(* IEC 61131-3 sources: daoli-st-library/DL_Device (part 36) *)

(* ---- FB_DL_VfdCapAgingEst.st ---- *)
(*
  ==================================================================
  组件名 Component  : FB_DL_VfdCapAgingEst
  分类   Category   : DL_Device
  前缀   Naming     : FB_DL_ ｜ b/n/u/f/t/e/st 类型前缀制（R265）
  码位   Code ID    : 16#0003_0725（故障级）｜ 16#0003_0726（信息级）
  版本   Version    : 1.0.0
  复杂度 Complexity  : 中
  功能   Purpose    : 母线电容老化趋势估计：纹波率实测值相对投运基线的长期比值监视
                      （电解电容容值衰减 → 纹波率单调爬升的运维预警）。
  开源溯源 Origin    : 公开公式 clean-room，参考公开电力电子运维工程口径的电解电容
                      纹波率基线比值判据（分类与公式借鉴，零代码复制），本件实现、
                      闸门与码位 100% 自有。
  许可证 License    : MIT
  参考   Reference  : IEC 61131-3:2013 §6.6 算术运算符；纹波率基线比值公开工程定义
  平台   Platform   : 纯 IEC 61131-3（四则 / 比较），三平台通用
  依赖   Depends    : 仅 Standard.library（无库调用、无定时器）
  分工声明 Split     : FB_DL_VfdDcBusRipple（瞬时纹波，R63 返修件）/ FB_DL_Brake
                      ResistorThermal（制动热）/ FB_DL_VfdThermalDerate（降额策略）
                      互引；本件为长期老化趋势，MANUAL 写明「瞬时监视与趋势估计
                      分层使用」（R216）。本件不实例依赖 VfdDcBusRipple，只收数值。
  归属 Ownership     : 本件无 TYPE 声明；全部引脚为 IEC 标准原生类型。
  ------------------------------------------------------------------
  边界 Boundary     :
                      一 组态闸结构早退（族② 判据，R1 同族教训出厂即正确）：
                         fRippleBasePct ≤ 0 或非有限（除子直穿防线）、fAgingLimPct ≤ 0
                         或非有限、fHystPct < 0 或非有限 → 组态码 0725 + 三件套 +
                         RETURN（除法段结构性不可达）；
                      二 fRipplePct 非有限或 < 0 → 该拍拒绝：比值冻结、迟滞态保持、
                         bValid = FALSE（丢弃 + 局部信息级计数，不外显 R62-D7 口径，
                         不影响趋势判据，禁污染物进除法）；
                      三 判据（带迟滞，两方向分别定义 R146）：fRippleRatioPct >
                         100 + fAgingLimPct 触发 bAgingHigh，回落 <
                         100 + fAgingLimPct×(1−fHystPct/100) 复原；
                      四 除子 fRippleBasePct > 0 已由段 2 结构早退证明（禁除零）；
                      五 负载可比性声明（写死）：本件假设同负载段比较，负载段切换时
                         调用方应 bEnable 短暂断开复位迟滞态——本件不自动判负载
                         （保持单一职责）；
                      六 bEnable = FALSE 的语义写死（FB33-4 声明行）：bAgingHigh 复位
                         + 比值冻结（运维趋势件，不丢历史）；
                      七 首拍 _bInit 全量初始化；无状态机（CASE N/A，R6 标注）；无
                         定时器 / 无边沿实例（段 0 无刷新对象）；无全局、无外部变量、
                         无物理地址、无指针。
  错误码 Codes      :
    16#0003_0725【故障级】组态非法（基线 ≤ 0 / 非有限；劣化阈值 ≤ 0 / 非有限；
                         迟滞 < 0 / 非有限）
    16#0003_0726【信息级】老化超限（bAgingHigh = TRUE，基线比超过 100 + 劣化阈值）
  码位反证 Note     :
    仅两码：0725 组态族为即刻判（与测点无关），0726 需比值已建立，处置人不同
    （组态工程师 / 运维），可由场景还原（R90）；fRipplePct 非有限拒绝拍不占码
    （bValid = FALSE 已足够表达，无额外处置信息，R90 不加码）。
  验收 Acceptance   :
    算法已证（脚本）：未跑 ｜ 编译器已证（三平台）：未跑
    V1 fRipplePct = fRippleBasePct → 比值 100%、bAgingHigh = FALSE
    V2 比值爬到 151%（限 150%）→ 触发；V3 回落 148%（迟滞未满足）→ 保持触发
    V4 回落 142% → 复原；V5 fRippleBasePct = 0 → 组态早退（R1 同族回归向量）
    V6 fRippleBasePct = NaN → 组态早退；V7 fRipplePct = NaN → 该拍拒绝不触发
    V8 fAgingLimPct = 0 → 组态早退（判据永假）
  修订记录 Revision  :
    2026-11-21  v1.0.0  R63 首版（批 4 · 序号 12）
  ==================================================================
*)
FUNCTION_BLOCK FB_DL_VfdCapAgingEst
VAR_INPUT
    bEnable       : BOOL := TRUE;  // 使能，FALSE 时判据复位 + 比值冻结（边界六）/ the enable, false resets the criterion and freezes the ratio
    fRipplePct    : LREAL := 0.0;  // 纹波率实测 [%]，由 FB_DL_VfdDcBusRipple 出口注入 / the measured ripple rate injected from the ripple monitor
    fRippleBasePct: LREAL := 5.0;  // 投运基线纹波率 [%]，须 > 0（除子）/ the commissioned baseline ripple rate, must be positive
    fAgingLimPct  : LREAL := 50.0; // 劣化阈值 [−]，相对基线百分比（50 即 150% 判劣化）/ the aging threshold relative to the baseline
    fHystPct      : LREAL := 5.0;  // 判据迟滞 [%]，须 ≥ 0 / the criterion hysteresis in percent, non negative
END_VAR
VAR_OUTPUT
    fRippleRatioPct : LREAL := 0.0;           // 基线比 fRipplePct/fRippleBasePct×100 [%] / the baseline ratio in percent
    bAgingHigh      : BOOL := FALSE;          // 老化超限判据（带迟滞）[-] / the aging high criterion with hysteresis
    bValid          : BOOL := FALSE;          // 判据可用 [-] / the criterion is usable
    eErr            : UDINT := 16#0000_0000;  // 错误码，0 = 正常 / the error code, zero is ok
    bError          : BOOL := FALSE;          // 故障标志（故障级码同拍置位，R45 配对）/ the fault flag raised with a fault level code
END_VAR
VAR
    _bInit      : BOOL := FALSE;   // 首拍初始化标志（R310 / FB50-2）/ the first scan flag
    _fRatio     : LREAL := 0.0;    // 基线比工作副本 [%] / the working baseline ratio
    _fRatioLast : LREAL := 0.0;    // 最近有效基线比（冻结源）[%] / the last valid ratio used while frozen
    _fTripLim   : LREAL := 0.0;    // 置警阈值 = 100 + 劣化阈值 [%] / the trip threshold
    _fReleLim   : LREAL := 0.0;    // 复原阈值 = 100 + 劣化阈值×(1−h) [%] / the release threshold
    _bAgingL    : BOOL := FALSE;   // 老化迟滞状态（跨拍保持）/ the aging hysteresis state
    _bFinBase   : BOOL := FALSE;   // 基线有限闸结果（逐拍重算）/ the baseline finiteness gate result
    _bFinLim    : BOOL := FALSE;   // 劣化阈值有限闸结果（逐拍重算）/ the threshold finiteness gate result
    _bFinHyst   : BOOL := FALSE;   // 迟滞有限闸结果（逐拍重算）/ the hysteresis finiteness gate result
    _bFinMeas   : BOOL := FALSE;   // 实测值有限闸结果（逐拍重算）/ the measurement finiteness gate result
    _bCfgBad    : BOOL := FALSE;   // 组态非法标记（逐拍重算）/ the configuration fault flag
    _nRejectCnt : DINT := 0;       // 实测值拒绝计数 [个]（仅局部留档，不外显，R62-D7 口径）/ the rejected measurement count, local only and never exposed
END_VAR  // R64 结构补齐：VAR 段缺失的 END_VAR（门禁机械修复）
VAR CONSTANT
    DL_VCA_PCT   : LREAL := 100.0; // 百分比换算与基线常量 [%] / the percentage scaling and the baseline constant
    DL_VCA_ZERO  : LREAL := 0.0;   // 实数零常量 [%] / the real zero constant
    DL_VCA_ONEI  : DINT := 1;      // 整型一常量 [个] / the integer one constant
    DL_VCA_ZEROI : DINT := 0;      // 整型零常量 [个] / the integer zero constant
END_VAR

// 段 0｜本件无定时器与边沿实例（纯趋势监视器，R6 标注 N/A），无刷新对象 / segment 0, no timers and no edge instances exist here

// 段 1｜首拍初始化（FB50-2）/ segment 1, the first scan init
IF NOT _bInit THEN // 首拍一拍 / the first scan
    _bInit := TRUE; // 置首拍标志 / raise the first scan flag
    _bAgingL := FALSE; // 迟滞态显式清零 / clear the hysteresis state explicitly
    _fRatioLast := DL_VCA_PCT; // 最近有效基线比显式预置 100%（首次有效计算前的安全占位）/ preset the last valid ratio to one hundred percent
    _nRejectCnt := DL_VCA_ZEROI; // 拒绝计数显式清零 [个] / clear the reject count explicitly
END_IF

// 段 2｜组态域闸结构早退（边界一，族② 判据：除子直穿防线先行，R272 全量点名）/ segment 2, the structural early exit on an illegal configuration
_bFinBase := (fRippleBasePct = fRippleBasePct) AND ((fRippleBasePct - fRippleBasePct) = (fRippleBasePct - fRippleBasePct)); // 基线有限 / the baseline is finite
_bFinLim := (fAgingLimPct = fAgingLimPct) AND ((fAgingLimPct - fAgingLimPct) = (fAgingLimPct - fAgingLimPct)); // 劣化阈值有限 / the threshold is finite
_bFinHyst := (fHystPct = fHystPct) AND ((fHystPct - fHystPct) = (fHystPct - fHystPct)); // 迟滞有限 / the hysteresis is finite
_bCfgBad := (NOT _bFinBase) OR (fRippleBasePct <= DL_VCA_ZERO)
         OR (NOT _bFinLim) OR (fAgingLimPct <= DL_VCA_ZERO)
         OR (NOT _bFinHyst) OR (fHystPct < DL_VCA_ZERO); // 组态非法 / an illegal configuration
IF _bCfgBad THEN // 组态非法：结构早退（出口三件套 + RETURN，除法段不可达）/ an illegal configuration exits structurally
    fRippleRatioPct := _fRatioLast; // 比值冻结最近有效值 [%]（禁自赋值出口，R261）/ freeze the last valid ratio
    bAgingHigh := FALSE; // 判据复位 / the criterion resets
    bValid := FALSE; // 判据不可用 / the criterion is not usable
    eErr := 16#0003_0725; // 故障级：组态非法 / fault grade, an illegal configuration
    bError := TRUE; // 同拍置故障标志（R45 配对）/ raise the fault flag on the same scan
    RETURN; // 结构早退 / the structural early exit
END_IF

// 段 3｜失能分支：判据复位 + 比值冻结（边界六声明行）/ segment 3, the disabled branch
IF NOT bEnable THEN // 失能 / disabled
    fRippleRatioPct := _fRatioLast; // 比值冻结最近有效值 [%]（运维趋势件，不丢历史）/ freeze the last valid ratio
    bAgingHigh := FALSE; // 判据复位 / the criterion resets
    bValid := FALSE; // 失能即不可用 / the criterion is not usable while disabled
    bError := FALSE; // 失能不是故障 / a disabled device is not a fault
    eErr := 16#0000_0000; // 失能不发码 / no code is emitted while disabled
    RETURN; // 早退 / early return
END_IF

// 段 4｜实测值拒绝闸（边界二：非有限或负值拒绝，禁污染物进除法）/ segment 4, the measurement rejection gate
_bFinMeas := (fRipplePct = fRipplePct) AND ((fRipplePct - fRipplePct) = (fRipplePct - fRipplePct)); // 实测值有限 / the measurement is finite
IF (NOT _bFinMeas) OR (fRipplePct < DL_VCA_ZERO) THEN // 实测坏或负值 / a broken or a negative measurement
    _nRejectCnt := _nRejectCnt + DL_VCA_ONEI; // 拒绝计数推进（仅局部留档，不外显）/ advance the reject count, local only
    fRippleRatioPct := _fRatioLast; // 比值冻结 [%] / freeze the ratio
    bAgingHigh := _bAgingL; // 迟滞态保持（拒绝拍不影响趋势判据）/ keep the hysteresis state
    bValid := FALSE; // 该拍不可用 / the scan is not usable
    eErr := 16#0000_0000; // 拒绝拍不发码（bValid = FALSE 已足够表达，R90 不加码）/ no code for a rejected scan
    bError := FALSE; // 无故障 / no fault
    RETURN; // 早退，除法不可达 / early return, the division is unreachable
END_IF

// 段 5｜基线比计算（除子 fRippleBasePct > 0 已由段 2 证明，禁除零）/ segment 5, the baseline ratio computation
_fRatio := (fRipplePct / fRippleBasePct) * DL_VCA_PCT; // 基线比 [%]，除子已证 > 0 / the baseline ratio with the proven divisor
_fRatioLast := _fRatio; // 最近有效基线比快照 [%] / snapshot the valid ratio
_fTripLim := DL_VCA_PCT + fAgingLimPct; // 置警阈值 [%] / the trip threshold
_fReleLim := DL_VCA_PCT + (fAgingLimPct * ((DL_VCA_PCT - fHystPct) / DL_VCA_PCT)); // 复原阈值 [%] / the release threshold

// 段 6｜老化判据迟滞（边界三，两方向分别定义，R146）/ segment 6, the aging hysteresis
IF NOT _bAgingL THEN // 未报警态 / the released state
    IF _fRatio > _fTripLim THEN // 超过置警阈值 / above the trip threshold
        _bAgingL := TRUE; // 置迟滞状态 / set the hysteresis state
    END_IF
ELSE // 已报警态 / the tripped state
    IF _fRatio < _fReleLim THEN // 回落低于复原阈值 / below the release threshold
        _bAgingL := FALSE; // 复原 / release
    END_IF
END_IF

// 段 7｜统一出口（迟滞状态派生，R187 / FB51-8）/ segment 7, the unified outlet
fRippleRatioPct := _fRatio; // 基线比出口 [%] / the ratio outlet
bAgingHigh := _bAgingL; // 判据出口 / the criterion outlet
bValid := TRUE; // 判据可用 / the criterion is usable
bError := FALSE; // 无故障 / no fault
IF _bAgingL THEN // 老化超限（信息级）/ the aging is high, informational
    eErr := 16#0003_0726; // 信息级：基线比超过 100 + 劣化阈值 / informational, the ratio exceeds the aging threshold
ELSE // 无事件 / no event
    eErr := 16#0000_0000; // 正常 / ok
END_IF
END_FUNCTION_BLOCK

(* ---- FB_DL_VfdCtrlWordBuild.st ---- *)
(*
  道莅工业代码库 | DL_Device | FB_DL_VfdCtrlWordBuild
  版本: 1.0.0 | 日期: 2026-11-23 | 轮次: R75
  开源溯源: brOscatLib (github.com/brOscatLib) / MIT / 借鉴 CtrlWordBuild 的语义，代码为 clean-room 重写
  功能: 变频器控制字编码——目标状态号（bit0..3）+ 命令位（运行/自由停车/直流
        制动/快速停止/反转/复位脉冲）按固定位图组装控制字；与 FB_DL_VfdStateWordMatch
        成对（编码/判码）。变换型 FB：无相位机，每拍独立全量重算。
  兼容性: CODESYS 3.5 / TwinCAT 3 / 汇川 InoProShop；仅依赖标准 R_TRIG，零厂商私有库
  接口: 输入 bEn/uStateNo（0..15，越界钳 15 并置信息码）/六命令位；输出
        wCtrlWord/uStateEff（钳位后状态号）/bRangeInfo/bError/nErrId。
  位图定义（bit0..3 = 目标状态号，与 C04 判码件低 4 位状态号口径一致）:
    bit4 = 运行命令 bRunCmd            bit5 = 非自由停车（1=斜坡停车可用）
    bit6 = 直流制动 bDCBrake           bit7 = 复位脉冲（R_TRIG 单拍）
    bit11 = 反转 bReverse              bit13 = 快速停止 bQuickStop
  码表: 16#0003_040F 信息级：目标状态号越域钳 15（每拍重算，非锁存）
        码段说明：0003 段信息子带 04xx，槽位经全库实扫空闲。
  边界: ① uStateNo > 15 → 钳 15 + bRangeInfo（本件无故障级路径，bError 恒 FALSE）；
        ② bit7 复位脉冲由 R_TRIG 单拍化（不复位脉冲不驻留控制字）；
        ③ bEn = FALSE 时控制字输出 16#0000（全零安全侧）；
        ④ R_TRIG 段 0 无条件周期刷新；⑤ 零全局耦合。
  邻件比对: StatusWordSegDecoder（通用分段译码 vs 本件变频器控制字编码组装）。
  修订历史: 2026-11-23 v1.0.0 R75 首版（复杂件批 B2 · C10）
*)

FUNCTION_BLOCK FB_DL_VfdCtrlWordBuild
VAR_INPUT
    bEn         : BOOL := FALSE;    // 编码使能（FALSE 输出全零控制字）[-] | Build enable, FALSE outputs zero word
    uStateNo    : UINT := 0;        // 目标状态号，域 [0, 15]，越界钳 15 [号] | Target state number, clamped to 15
    bRunCmd     : BOOL := FALSE;    // 运行命令（bit4）[-] | Run command bit
    bCoastStop  : BOOL := FALSE;    // 自由停车选择（TRUE 时 bit5=0）[-] | Coast stop select, TRUE clears bit5
    bDCBrake    : BOOL := FALSE;    // 直流制动（bit6）[-] | DC brake bit
    bQuickStop  : BOOL := FALSE;    // 快速停止（bit13）[-] | Quick stop bit
    bReverse    : BOOL := FALSE;    // 反转（bit11）[-] | Reverse bit
    bResetCmd   : BOOL := FALSE;    // 故障复位命令（bit7，沿触发单拍）[-] | Fault reset command, edge one-shot
END_VAR
VAR_OUTPUT
    wCtrlWord  : WORD;              // 组装控制字出口（bEn=FALSE 时全零）[-] | Built control word outlet
    uStateEff  : UINT;              // 钳位后状态号出口 [号] | Clamped state number outlet
    bRangeInfo : BOOL;              // 状态号越域钳位当拍信息 [-] | Range clamp info this scan
    bError     : BOOL;              // 故障标志（本件无故障路径，恒 FALSE）[-] | Error flag, no fault paths
    nErrId     : UDINT;             // 事件码，0 = 无事件 | Event code, 0 = none
END_VAR
VAR
    _uStateEff : UINT := 0;         // 钳位状态号内部镜像 [号] | Clamped state number mirror
    _wOut      : WORD := 16#0000;   // 组装暂存字 [-] | Build staging word
    _bRange    : BOOL;              // 越域当拍量 [-] | Range violation this scan
    rtResetCmd : R_TRIG;            // 复位脉冲沿实例，段 0 无条件刷新 | Reset pulse edge instance
END_VAR

(* —— 段 0：沿实例无条件周期刷新（R7 红线） —— *)
rtResetCmd(CLK := bResetCmd);                 // 复位脉冲沿每拍必调 / Reset pulse edge every scan

(* —— 段 1：状态号钳位（越域置当拍信息量） —— *)
_uStateEff := uStateNo;                       // 状态号暂存 / State number staging
_bRange := FALSE;                             // 越域当拍量预清 / Range flag preset
IF _uStateEff > 15 THEN
    _uStateEff := 15;                         // 越域钳 15 / Clamp to 15
    _bRange := TRUE;                          // 置越域信息量 / Set range info
END_IF

(* —— 段 2：控制字位图组装（bit0..3 状态号） —— *)
_wOut := INT_TO_WORD(UINT_TO_INT(_uStateEff)) AND 16#000F;    // 状态号入低 4 位（掩码兜底）/ State number to low nibble
IF bRunCmd THEN
    _wOut := _wOut OR 16#0010;                // bit4 运行命令 / Run command bit
END_IF
IF NOT bCoastStop THEN
    _wOut := _wOut OR 16#0020;                // bit5 斜坡停车可用（非自由停车）/ Ramp stop available bit
END_IF
IF bDCBrake THEN
    _wOut := _wOut OR 16#0040;                // bit6 直流制动 / DC brake bit
END_IF
IF rtResetCmd.Q THEN
    _wOut := _wOut OR 16#0080;                // bit7 复位脉冲（仅沿当拍驻留）/ Reset pulse bit, one scan only
END_IF
IF bReverse THEN
    _wOut := _wOut OR 16#0800;                // bit11 反转 / Reverse bit
END_IF
IF bQuickStop THEN
    _wOut := _wOut OR 16#2000;                // bit13 快速停止 / Quick stop bit
END_IF

(* —— 段 3：出口单点映射（名实同源；信息码每拍重算） —— *)
IF bEn THEN
    wCtrlWord := _wOut;                       // 使能输出组装字 / Enabled, output built word
ELSE
    wCtrlWord := 16#0000;                     // 未使能输出全零（安全侧） / Disabled, output zero word
END_IF
uStateEff := _uStateEff;                      // 钳位状态号出口 / Clamped state outlet
bRangeInfo := _bRange;                        // 越域信息出口 / Range info outlet
bError := FALSE;                              // 本件无故障级路径（头注释声明）/ No fault paths by design
IF _bRange THEN
    nErrId := 16#0003_040F;                   // 信息级：状态号越域钳位 / Info: state number clamped
ELSE
    nErrId := 16#0000_0000;                   // 无事件 / No event
END_IF

END_FUNCTION_BLOCK

(* ---- FB_DL_VfdGeneric.st ---- *)
(*==============================================================================
 * 组件名称 (Component)  : FB_DL_VfdGeneric
 * 所属子库 (Sublibrary) : DL_Device
 * 当前版本 (Version)    : 1.0.1
 * 兼容性   (Platform)   : CODESYS 3.5 / TwinCAT 3 / 汇川 InoProShop / Machine Expert
 *                         仅依赖 Standard.library（TON / R_TRIG / TP），零厂商方言
 * 分类     (Category)   : 设备执行器功能块（Function Block，实现 I_DL_VfdDrive）
 * 功能简述 (Function)   : 通用变频器端子型控制功能块。正/反转端子互斥
 *                         （出口断言 + 冲突安全侧停止）、点动优先覆盖运行、
 *                         多段速表/模拟量给定双通道频率设定（越界钳位）、
 *                         频率给定模拟量域线性映射、指令-反馈校验窗、驱动
 *                         故障锁存与复位端子定宽脉冲重试；状态机
 *                         E_DL_VfdState + CASE + ELSE 兜底。
 * 接口实现 (Implements) : I_DL_VfdDrive。接口 OUT 列同名成员（eState/
 *                         fFreqSetpoint/fFreqActual/bRunning/bFault/
 *                         uErrorId）按 R22 以只读 PROPERTY GET 承载（内部
 *                         镜像同源），非接口成员 bRunFwdOut/bRunRevOut/
 *                         bJogOut/bFaultResetOut/fFreqRefPercent/uPresetCode
 *                         保留 VAR_OUTPUT；方法 CmdRun/CmdStop/CmdJog/
 *                         SetFrequency/SelectPresetSpeed/CmdReset 全部在
 *                         本文件尾部落地。
 * 开源溯源 (Origin)     : 来源标签 lbp-basic-process / lbp-device
 *                         （RAW_NOTES_R6 S-1 + S-4：变频器端子标准信号集
 *                         ——正反转互斥、点动优先、多段速 DI 组合、模拟
 *                         量频率给定线性映射、故障复位端子脉冲等行业公知
 *                         工程惯例，公开技术资料，仅借鉴通用信号域语义；
 *                         状态机、钳位与互斥实现、故障码按本库红线独立
 *                         设计，clean-room 未复制源码）。
 * 红线自检 (Redline)    : R1 零全局变量表/外部变量引用 ✓｜R2 零物理 IO 地址 ✓
 *                         R3 纯 IEC 61131-3 ✓｜R4 防除零/防越界/非有限值
 *                         防御/浮点容差比较 ✓｜R5 全变量中英双语同行注释 ✓
 *                         R6 ENUM+CASE+ELSE ✓｜R7 三个定时器/边缘/脉冲实例
 *                         主体最前部无条件刷新 ✓
 * 公约遵循 (Convention) : 0.1/R23 本块为纯事件型状态机（BOOL 指令/反馈 +
 *                         频率标量直通计算，无积分/滤波类连续量同步语义），
 *                         免首扫，无内部初始化标志。
 *                         0.7 故障码段位 16#0003_xxxx：【故障级】0003_0250
 *                         驱动故障 / 0003_0251 启动反馈超时 / 0003_0252
 *                         非法状态，R15 锁存仅复位脉冲路径可清；【信息级】
 *                         0003_0106 正反转指令冲突 / 0003_0107 频率设定
 *                         钳位/段速选择越界（瞬时型每拍重算，0.15）。
 * 偏离留档 (Deviation)  : 依 R11 头注释留档，共 2 条：
 *                         ① 信息级码：规格原分配 0003_0103/0104，经与子库
 *                           VERSION.md 故障码表核对，R5 已占用 0102~0104
 *                           （AnalogTransmitter），依公约 0.7 冲突顺延为
 *                           0003_0106/0107（0105 经终审裁定空置：重启抑制
 *                           拒绝统一沿用 DolMotor 既有语义码位 0003_0208，
 *                           见 FB_DL_StarDeltaMotor 终审记录）。
 *                         ② 点动频率：规格设计要点"点动频率取 aPresetFreq[1]
 *                           （注释声明）"落为引脚注释声明——本块不因点动切
 *                           换频率通道（端子型变频器点动频率由驱动器内部组
 *                           态承担），段速 1 兼作点动频率域供现场整定选用。
 * 修订历史 (Revision)   :
 *   2026-11-15  v1.0.0  首版入库（R6 轮 · DL_Device 阀门/驱动族深化）
 *   2026-11-15  v1.0.1  终审修复【致命】复位端子脉冲触发时序：原实现
 *                       _bResetPulseReq 于主体末尾同拍自清，TP 实例（段 1
 *                       最前部刷新）永远采不到 TRUE 入参，bFaultResetOut
 *                       恒 FALSE，故障复位端子脉冲永不输出（验收向量 V5
 *                       不成立，R13 逐拍推演复现）。修法：自清动作移至
 *                       TP 实例调用之后。另补点动频率引脚注释声明（R11
 *                       偏离②）。引脚契约零变更。
 *============================================================================*)
FUNCTION_BLOCK FB_DL_VfdGeneric IMPLEMENTS I_DL_VfdDrive
VAR_INPUT
    bDriveEnable     : BOOL;            // 驱动使能/上电（Drive enable），FALSE → 未使能态全部输出切断 / Drive enable, FALSE cuts off all outputs
    bCmdRunFwd       : BOOL;            // 正转运行指令（Run forward command），电平生效 / Run forward command, level effective
    bCmdRunRev       : BOOL;            // 反转运行指令（Run reverse command），电平生效；与正转同拍为真 → 冲突安全侧停止 / Run reverse command, conflict with forward stops safely
    bCmdJogFwd       : BOOL;            // 正向点动指令（Jog forward command），电平生效，优先级高于运行指令；点动频率不在本块内切换通道——端子型惯例由驱动器内部点动频率组态承担，亦可现场将 aPresetFreq[1] 整定为点动频率域（段速 1 兼作点动频率） / Jog forward command, level effective, priority over run; jog frequency not switched by this block, use drive-internal jog frequency or tune aPresetFreq[1] as the jog frequency domain
    bFbRunning       : BOOL;            // 运行反馈（Running feedback），TRUE=驱动输出运行中 / Running feedback, TRUE = drive output running
    bFbFault         : BOOL;            // 驱动故障反馈（Drive fault feedback），TRUE=故障 / Drive fault feedback, TRUE = faulty
    bFbAtSpeed       : BOOL;            // 频率到达反馈（At-speed feedback），TRUE=输出频率到达设定容差带 / At-speed feedback, TRUE = output frequency reached setpoint band
    fFreqCmd         : REAL;            // 频率设定（Frequency command）[Hz]，0..fFreqMax，越界钳位信息级 / Frequency command [Hz], clamped with info code
    fFreqActual      : REAL;            // 频率反馈（Frequency feedback）[Hz]，非有限值防御 / Frequency feedback [Hz], non-finite defended
    aPresetFreq      : ARRAY[1..7] OF REAL; // 多段速频率表（Preset speed table）[Hz]，段速值由现场整定注入 / Preset speed table [Hz], field-tuned values injected
    nPresetSel       : USINT;           // 段速选择（Preset speed select），0=模拟量给定、1..7=段速，越界按 0 处理并置码 / Preset select, 0 = analog reference, 1..7 = steps, out-of-range treated as 0 with code
    fFreqMax         : REAL := 50.0;    // 频率上限（Max frequency）[Hz]，默认 50.0 / Maximum frequency [Hz], default 50.0
    tFbWindow        : TIME := T#1S;    // 指令-反馈校验窗口（Feedback check window），T#0S=免校验 / Feedback check window, T#0S disables the check
    tFaultResetPulse : TIME := T#500MS; // 故障复位脉冲宽度（Fault reset pulse）/ Fault reset pulse width
    bReset           : BOOL;            // 故障复位请求（Fault reset request），上升沿生效 / Fault reset request, rising edge effective
END_VAR

VAR_OUTPUT
    bRunFwdOut      : BOOL;             // 正转端子输出（Run forward terminal）/ Run forward terminal output
    bRunRevOut      : BOOL;             // 反转端子输出（Run reverse terminal）/ Run reverse terminal output
    bJogOut         : BOOL;             // 点动端子输出（Jog terminal）/ Jog terminal output
    bFaultResetOut  : BOOL;             // 故障复位端子输出（Fault reset terminal），tFaultResetPulse 定宽单发 / Fault reset terminal, one-shot fixed-width pulse
    fFreqRefPercent : REAL;             // 频率给定模拟量输出（Frequency reference analog out）[%]，0~100 线性映射 fFreqMax / Analog frequency reference [%], linear over fFreqMax
    uPresetCode     : USINT;            // 段速选择码输出（Preset speed code），映射 DI 多段速端子组合 0..7 / Preset speed code mapped to DI terminal group 0..7
END_VAR

VAR
    _eState         : E_DL_VfdState := E_DL_VfdState.eDisabled; // 内部状态机步序（Internal state step），外部经属性只读 / Internal state, read-only via property
    _bFaultLatch    : BOOL;             // 故障锁存标志（Fault latch flag），仅复位脉冲路径清除 / Fault latch flag, cleared only via reset pulse path
    _uErrorIdInt    : UDINT;            // 内部故障码寄存（Internal error register），故障级与信息级共用 / Internal error register, fault and info codes share it
    _uInfoCode      : UDINT;            // 本拍信息级码（Info code this cycle），瞬时型每拍重算（0.15）/ Transient info code recomputed each cycle
    _bPendRunFwd    : BOOL;             // 方法正转保持锁存（Method run-forward hold latch）/ Method run-forward hold latch
    _bPendRunRev    : BOOL;             // 方法反转保持锁存（Method run-reverse hold latch）/ Method run-reverse hold latch
    _bJogHold       : BOOL;             // 方法点动保持锁存（Method jog hold latch）/ Method jog hold latch
    _bPendReset     : BOOL;             // 方法复位请求（Method reset request）/ Method reset request
    _bResetPulseReq : BOOL;             // 复位脉冲单拍触发请求（Reset pulse trigger request），置位一拍 / One-cycle reset pulse trigger request
    _fFreqMethodVal : REAL;             // 方法频率设定值（Method frequency value）[Hz] / Frequency value set via method
    _bFreqMethodAct : BOOL;             // 方法频率设定激活（Method frequency active），激活后覆盖引脚给定 / Method frequency active, overrides pin reference
    _uPresetMethod  : USINT;            // 方法段速选择值（Method preset select value）/ Preset select value set via method
    _bPresetMethodAct : BOOL;           // 方法段速选择激活（Method preset select active）/ Method preset select active flag
    _fFreqMaxEff    : REAL := 50.0;     // 防御后频率上限（Sanitized max frequency）[Hz] / Sanitized maximum frequency
    _fFreqCmdEff    : REAL := 0.0;      // 防御后模拟量给定（Sanitized analog command）[Hz]，非数回零 / Sanitized analog command, NaN falls back to zero
    _fFreqSetInt    : REAL := 0.0;      // 钳位后生效频率设定（Effective clamped setpoint）[Hz] / Effective clamped frequency setpoint
    _fFreqActHold   : REAL := 0.0;      // 末次有效频率反馈（Last valid frequency feedback）[Hz] / Last valid frequency feedback hold carrier
    _uPresetSelEff  : USINT;            // 钳位后生效段速选择（Effective clamped preset select），0..7 / Effective preset select clamped to 0..7
    _bRunFwd        : BOOL;             // 合成正转指令（Merged run-forward command），引脚 OR 方法锁存 / Merged forward command, pin OR method latch
    _bRunRev        : BOOL;             // 合成反转指令（Merged run-reverse command），引脚 OR 方法锁存 / Merged reverse command, pin OR method latch
    _bJog           : BOOL;             // 合成点动指令（Merged jog command），引脚 OR 方法锁存 / Merged jog command, pin OR method latch
    _bConflict      : BOOL;             // 正反转同拍冲突（Forward/reverse conflict this cycle）/ Forward-reverse conflict flag
    _bFbWinEn       : BOOL;             // 反馈校验窗使能（Feedback window enable），窗口参数大于零有效 / Feedback window enable, active when window above zero
    _bInFbWin       : BOOL;             // 反馈校验窗计时条件（Feedback window timing condition）/ Timing condition of feedback window
    _fbTrigReset    : R_TRIG;           // 引脚复位上升沿（Pin reset edge）/ Pin reset rising edge
    _fbTonFbWindow  : TON;              // 启动反馈校验窗定时器（Startup feedback window timer）/ Startup feedback window timer
    _fbTpResetPulse : TP;               // 复位端子定宽脉冲定时器（Reset terminal pulse timer），IEC 标准 TP / Reset terminal pulse timer, IEC standard TP
END_VAR

METHOD CmdRun : BOOL
VAR_INPUT
    bFwd : BOOL; // 方向选择（Direction select），TRUE=正转 / FALSE=反转 / TRUE = forward, FALSE = reverse
END_VAR
IF _bFaultLatch OR (_eState = E_DL_VfdState.eFault) OR (_eState = E_DL_VfdState.eDisabled) THEN
    CmdRun := FALSE;          // 故障/未使能态拒绝（Rejected in fault or disabled state）
ELSE
    IF bFwd THEN
        _bPendRunFwd := TRUE; // 登记正转保持锁存（Register forward hold latch）
        _bPendRunRev := FALSE; // 互斥注销反转锁存（Cancel opposite latch）
    ELSE
        _bPendRunRev := TRUE; // 登记反转保持锁存（Register reverse hold latch）
        _bPendRunFwd := FALSE; // 互斥注销正转锁存（Cancel opposite latch）
    END_IF
    CmdRun := TRUE;           // 受理成功（Accepted）
END_IF

(*------------------------------------------------------------------------------
 * 方法: CmdStop —— 停止指令：撤销运行/点动锁存，无条件受理。
 *      Method CmdStop - revokes run and jog latches, unconditionally accepted.
 *------------------------------------------------------------------------------*)
    END_METHOD

METHOD CmdStop : BOOL
VAR_INPUT
END_VAR
_bPendRunFwd := FALSE;        // 撤销正转锁存（Release forward latch）
_bPendRunRev := FALSE;        // 撤销反转锁存（Release reverse latch）
_bJogHold    := FALSE;        // 撤销点动保持（Release jog hold）
CmdStop := TRUE;              // 无条件受理（Unconditionally accepted）

(*------------------------------------------------------------------------------
 * 方法: CmdJog —— 点动指令（bFwd=TRUE 登记保持 / FALSE 撤销）。故障态拒绝。
 *      Method CmdJog - jog hold register/release, rejected in fault state.
 *------------------------------------------------------------------------------*)
    END_METHOD

METHOD CmdJog : BOOL
VAR_INPUT
    bFwd : BOOL; // 点动方向（Jog direction），TRUE=正向登记 / FALSE=撤销保持 / TRUE = register, FALSE = release
END_VAR
IF _bFaultLatch OR (_eState = E_DL_VfdState.eFault) THEN
    CmdJog := FALSE;          // 故障态拒绝（Rejected in fault state）
ELSE
    _bJogHold := bFwd;        // 登记或撤销点动保持（Register or release jog hold）
    CmdJog := TRUE;           // 受理成功（Accepted）
END_IF

(*------------------------------------------------------------------------------
 * 方法: SetFrequency —— 频率设定 [Hz]，越界/非有限值拒绝返回 FALSE。
 *      Method SetFrequency - frequency set, out-of-range or NaN returns FALSE.
 *------------------------------------------------------------------------------*)
    END_METHOD

METHOD SetFrequency : BOOL
VAR_INPUT
    fHz : REAL; // 频率设定值（Frequency value）[Hz]，域 0..fFreqMax / Frequency value [Hz], range 0..fFreqMax
END_VAR
IF (fHz <> fHz) OR (fHz < 0.0) OR (fHz > _fFreqMaxEff) THEN
    SetFrequency := FALSE;    // 非数或越域拒绝（Rejected on NaN or out of range）
ELSE
    _fFreqMethodVal := fHz;   // 登记方法频率设定（Register method frequency value）
    _bFreqMethodAct := TRUE;  // 激活方法给定通道（Activate method reference channel）
    SetFrequency := TRUE;     // 受理成功（Accepted）
END_IF

(*------------------------------------------------------------------------------
 * 方法: SelectPresetSpeed —— 多段速选择，0=模拟量给定、1..7=段速，越界拒绝。
 *      Method SelectPresetSpeed - preset select, 0 = analog, 1..7 = steps.
 *------------------------------------------------------------------------------*)
    END_METHOD

METHOD SelectPresetSpeed : BOOL
VAR_INPUT
    nIdx : USINT; // 段速索引（Preset index），0=模拟量给定 / 1..7=段速 / Preset index, 0 = analog reference, 1..7 = steps
END_VAR
IF nIdx <= 7 THEN
    _uPresetMethod := nIdx;   // 登记方法段速选择（Register method preset value）
    _bPresetMethodAct := TRUE; // 激活方法段速通道（Activate method preset channel）
    SelectPresetSpeed := TRUE; // 受理成功（Accepted）
ELSE
    SelectPresetSpeed := FALSE; // 越界拒绝（Rejected on out-of-range index）
END_IF

(*------------------------------------------------------------------------------
 * 方法: CmdReset —— 复位指令，返回是否受理（存在锁存故障时为 TRUE）。
 *      Method CmdReset - reset command, returns TRUE only when latch exists.
 *------------------------------------------------------------------------------*)
    END_METHOD

METHOD CmdReset : BOOL
VAR_INPUT
END_VAR
IF _bFaultLatch OR (_eState = E_DL_VfdState.eFault) THEN
    _bPendReset := TRUE;      // 登记复位请求，主体状态机消化（Register reset request, consumed by body）
    CmdReset := TRUE;         // 可复位（Resettable）
ELSE
    CmdReset := FALSE;        // 无故障可复位（Nothing to reset）
END_IF

(*------------------------------------------------------------------------------
 * 属性: eState（GET）—— 当前状态机状态只读视图。
 *      Property eState (GET) - read-only view of the current state machine state.
 *------------------------------------------------------------------------------*)
    END_METHOD

// ============================================================================
// 段 1｜定时器与边缘检测实例无条件周期刷新（R7：严禁置于 IF/CASE 分支内）
//      Unconditional per-cycle refresh of all timer and edge instances (R7)
// ============================================================================
_fbTrigReset(CLK := bReset);
_bFbWinEn := (tFbWindow > T#0S);      // 窗口为零 = 免校验（Zero window = check disabled）
_bInFbWin := ((_eState = E_DL_VfdState.eRunningFwd) OR (_eState = E_DL_VfdState.eRunningRev))
             AND (NOT bFbRunning) AND _bFbWinEn; // 运行态且反馈未到才计时（Timing only while running and feedback pending）
_fbTonFbWindow(IN := _bInFbWin, PT := tFbWindow);
_fbTpResetPulse(IN := _bResetPulseReq, PT := tFaultResetPulse); // 复位端子定宽脉冲（Fixed-width reset terminal pulse）
_bResetPulseReq := FALSE;             // 单拍触发请求在 TP 采样后立即自清：TP 于本拍见到
                                      // TRUE 并起振，下一拍入参回落 FALSE，定宽由 TP 保持
                                      // （One-cycle trigger cleared right after TP sampling）

// ============================================================================
// 段 2｜参数防御（0.8：非数自比检测，默认值先赋）+ 指令合成与钳位
//      Parameter sanitation (0.8 NaN self-compare) + command merge and clamping
// ============================================================================
_uInfoCode := 0;                      // 本拍信息级码先归零，事件段重算（Info code preset zero, recomputed in event chain）
_fFreqMaxEff := fFreqMax;             // 频率上限镜像（Max frequency mirror）
IF _fFreqMaxEff <> _fFreqMaxEff THEN  // 非数自比检测（NaN self-compare test）
    _fFreqMaxEff := 50.0;             // 回落默认上限（Fallback to default max）
END_IF
IF ABS(_fFreqMaxEff) < 1E-6 THEN
    _fFreqMaxEff := 1E-6;             // 防除零：上限退化时钳最小正值（Divide-by-zero guard, degenerate max clamped to tiny positive）
END_IF

IF _bFreqMethodAct THEN
    _fFreqCmdEff := _fFreqMethodVal;  // 方法设定覆盖引脚给定（Method value overrides pin reference）
ELSE
    _fFreqCmdEff := fFreqCmd;         // 引脚模拟量给定（Pin analog reference）
END_IF
IF _fFreqCmdEff <> _fFreqCmdEff THEN  // 非数自比检测（NaN self-compare test）
    _fFreqCmdEff := 0.0;              // 非数给定回零（NaN reference falls back to zero）
END_IF
IF _fFreqCmdEff < 0.0 THEN
    _fFreqCmdEff := 0.0;              // 负给定下限钳位（Negative reference clamped to zero）
    _uInfoCode := 16#0003_0107;       // 0003_0107 频率设定钳位【信息级】/ Frequency clamped, info level
END_IF
IF _fFreqCmdEff > _fFreqMaxEff THEN
    _fFreqCmdEff := _fFreqMaxEff;     // 超上限钳位（Reference clamped to max）
    _uInfoCode := 16#0003_0107;       // 0003_0107 频率设定钳位【信息级】/ Frequency clamped, info level
END_IF

IF fFreqActual = fFreqActual THEN     // 频率反馈有效性（Frequency feedback validity）
    _fFreqActHold := fFreqActual;     // 更新末次有效反馈（Update last valid feedback）
END_IF                                 // 非有限值保持末次有效值（Non-finite holds last valid）

// 段速选择钳位：越界按 0 处理并置码（Preset select clamped, out-of-range as 0 with code）
IF _bPresetMethodAct THEN
    _uPresetSelEff := _uPresetMethod; // 方法段速选择覆盖引脚（Method preset overrides pin）
ELSIF nPresetSel <= 7 THEN
    _uPresetSelEff := nPresetSel;     // 引脚段速选择合法（Pin preset select valid）
ELSE
    _uPresetSelEff := 0;              // 越界按模拟量给定处理（Out-of-range treated as analog reference）
    _uInfoCode := 16#0003_0107;       // 0003_0107 段速选择越界【信息级】/ Preset select out of range, info level
END_IF

// 生效频率设定：段速优先，模拟量给定兜底（Effective setpoint: preset first, analog fallback）
IF (_uPresetSelEff >= 1) AND (_uPresetSelEff <= 7) THEN
    _fFreqSetInt := aPresetFreq[_uPresetSelEff];       // 取段速表值（Take preset table value, index proven 1..7）
    IF _fFreqSetInt <> _fFreqSetInt THEN
        _fFreqSetInt := 0.0;                           // 段速值非数回零防御（NaN preset falls back to zero）
    END_IF
ELSE
    _fFreqSetInt := _fFreqCmdEff;     // 模拟量给定通道（Analog reference channel）
END_IF

// 指令合成与冲突判定（Command merge and conflict evaluation）
_bRunFwd := bCmdRunFwd OR _bPendRunFwd; // 合成正转（Merged forward）
_bRunRev := bCmdRunRev OR _bPendRunRev; // 合成反转（Merged reverse）
_bJog := bCmdJogFwd OR _bJogHold;       // 合成点动，优先级最高（Merged jog, highest priority）
_bConflict := _bRunFwd AND _bRunRev;    // 同拍正反转冲突（Same-cycle conflict）
IF _bConflict THEN
    _uInfoCode := 16#0003_0106;         // 0003_0106 正反转指令冲突【信息级】/ Forward-reverse conflict, info level
END_IF

// ============================================================================
// 段 3｜驱动故障全局监视（优先级最高）：故障反馈置锁存
//      Drive fault global monitor (highest priority): fault feedback latches
// ============================================================================
IF bFbFault THEN
    _bFaultLatch := TRUE;               // 驱动故障锁存（Drive fault latch）
    _uErrorIdInt := 16#0003_0250;       // 0003_0250 驱动故障【故障级】/ Drive fault, fault level
    _eState      := E_DL_VfdState.eFault; // 强制故障态（Force fault state）
ELSIF (_eState = E_DL_VfdState.eRunningFwd) OR (_eState = E_DL_VfdState.eRunningRev) THEN
    IF _bFbWinEn AND _fbTonFbWindow.Q AND (NOT bFbRunning) THEN
        _bFaultLatch := TRUE;           // 启动反馈超时锁存（Startup feedback timeout latch）
        _uErrorIdInt := 16#0003_0251;   // 0003_0251 启动反馈超时【故障级】/ Startup feedback timeout, fault level
        _eState      := E_DL_VfdState.eFault;
    END_IF
END_IF

// ============================================================================
// 段 4｜核心状态机（ENUM + CASE，含 ELSE 非法状态兜底）
//      Core state machine (ENUM + CASE with ELSE illegal-state fallback)
// ============================================================================
IF _bFaultLatch OR (_eState = E_DL_VfdState.eFault) THEN
    CASE _eState OF
        E_DL_VfdState.eFault: // 故障锁存态：复位端子定宽脉冲重试恢复
            IF _bPendReset OR _fbTrigReset.Q THEN
                _bResetPulseReq := TRUE;        // 触发复位端子脉冲（Trigger reset terminal pulse）
                _bPendReset     := FALSE;       // 消费复位请求（Consume reset request）
                IF NOT bFbFault THEN
                    _bFaultLatch := FALSE;      // 驱动故障已消失，解除锁存（Drive fault cleared, release latch）
                    _uErrorIdInt := 0;          // 故障码清零（Error code cleared）
                    _eState      := E_DL_VfdState.eReady; // 回就绪态（Back to ready）
                END_IF
            END_IF
        ELSE // 锁存标志与状态不一致兜底：强制同步进故障态（Latch/state mismatch fallback）
            _eState := E_DL_VfdState.eFault;
    END_CASE
ELSIF NOT bDriveEnable THEN
    _eState     := E_DL_VfdState.eDisabled; // 未使能态：全部输出切断（Disabled: all outputs cut off）
    _bJogHold   := FALSE;                   // 撤销点动保持（Release jog hold）
    _bPendRunFwd := FALSE;                  // 撤销方法运行锁存（Release method run latches）
    _bPendRunRev := FALSE;
ELSE
    CASE _eState OF

        E_DL_VfdState.eDisabled: // 未使能态：等待使能
            _eState := E_DL_VfdState.eReady; // 使能完成转就绪（Enabled, to ready）

        E_DL_VfdState.eReady: // 就绪态：评估点动/运行指令
            IF _bJog THEN
                _eState := E_DL_VfdState.eJogging; // 点动优先受理（Jog accepted with priority）
            ELSIF _bConflict THEN
                // 正反转同拍冲突：安全侧保持停止（Conflict: hold safe-side stop）
            ELSIF _bRunFwd THEN
                _eState := E_DL_VfdState.eRunningFwd; // 正转受理（Forward accepted）
            ELSIF _bRunRev THEN
                _eState := E_DL_VfdState.eRunningRev; // 反转受理（Reverse accepted）
            END_IF

        E_DL_VfdState.eRunningFwd: // 正转运行态
            IF _bJog THEN
                _eState := E_DL_VfdState.eJogging; // 点动覆盖运行（Jog overrides run）
            ELSIF _bConflict OR (NOT _bRunFwd) THEN
                _eState := E_DL_VfdState.eReady;   // 冲突或指令撤销：安全侧回就绪（Conflict or command dropped: safe-side to ready）
            END_IF

        E_DL_VfdState.eRunningRev: // 反转运行态
            IF _bJog THEN
                _eState := E_DL_VfdState.eJogging; // 点动覆盖运行（Jog overrides run）
            ELSIF _bConflict OR (NOT _bRunRev) THEN
                _eState := E_DL_VfdState.eReady;   // 冲突或指令撤销：安全侧回就绪（Conflict or command dropped: safe-side to ready）
            END_IF

        E_DL_VfdState.eJogging: // 点动态：点动电平维持
            IF NOT _bJog THEN
                IF _bConflict THEN
                    _eState := E_DL_VfdState.eReady;             // 冲突安全侧回就绪（Conflict: safe-side to ready）
                ELSIF _bRunFwd THEN
                    _eState := E_DL_VfdState.eRunningFwd;        // 点动结束回正转（Jog ended, back to forward）
                ELSIF _bRunRev THEN
                    _eState := E_DL_VfdState.eRunningRev;        // 点动结束回反转（Jog ended, back to reverse）
                ELSE
                    _eState := E_DL_VfdState.eReady;             // 点动结束回就绪（Jog ended, back to ready）
                END_IF
            END_IF

        ELSE // 非法状态兜底：任何越界枚举值强制锁存故障（Illegal state fallback）
            _bFaultLatch := TRUE;                // 故障锁存（Fault latched）
            _uErrorIdInt := 16#0003_0252;        // 0003_0252 非法状态【故障级】/ Illegal state, fault level
            _eState      := E_DL_VfdState.eFault;
    END_CASE
END_IF

// ============================================================================
// 段 5｜输出推导 + 正/反转端子互斥出口断言（硬约束：两端子恒不可同真）
//      Output derivation + forward/reverse terminal exclusivity exit assertion
// ============================================================================
bRunFwdOut := (_eState = E_DL_VfdState.eRunningFwd); // 正转端子随状态（Forward terminal follows state）
bRunRevOut := (_eState = E_DL_VfdState.eRunningRev); // 反转端子随状态（Reverse terminal follows state）
bJogOut    := (_eState = E_DL_VfdState.eJogging);    // 点动端子随状态（Jog terminal follows state）
IF bRunFwdOut AND bRunRevOut THEN
    bRunFwdOut := FALSE;                  // 断言对调：异常同真时双断保安全（Assertion fallback: cut both on impossible condition）
    bRunRevOut := FALSE;
    _eState    := E_DL_VfdState.eReady;   // 强制回就绪（Force back to ready）
END_IF
IF (_eState = E_DL_VfdState.eDisabled) OR (_eState = E_DL_VfdState.eFault) THEN
    bRunFwdOut := FALSE;                  // 未使能/故障态全端子必断（Assertion: terminals off in disabled/fault）
    bRunRevOut := FALSE;
    bJogOut    := FALSE;
END_IF
bFaultResetOut := _fbTpResetPulse.Q;      // 复位端子定宽脉冲输出（Reset terminal pulse output）
uPresetCode := _uPresetSelEff;            // 段速码输出（Preset code output）
fFreqRefPercent := _fFreqCmdEff * (100.0 / _fFreqMaxEff); // 模拟量域线性映射，除数已证明非零（Linear analog mapping, divisor proven non-zero）

(*------------------------------------------------------------------------------
 * 方法: CmdRun —— 正/反转运行指令（受理为保持锁存）。故障/未使能态拒绝。
 *      Method CmdRun - run command held as latch, rejected in fault/disabled.
 *------------------------------------------------------------------------------*)

PROPERTY eState : E_DL_VfdState
eState := _eState;            // 返回内部状态（Return internal state）

(*------------------------------------------------------------------------------
 * 属性: fFreqSetpoint（GET）—— 钳位后生效频率设定 [Hz]。
 *      Property fFreqSetpoint (GET) - effective clamped frequency setpoint [Hz].
 *------------------------------------------------------------------------------*)
PROPERTY fFreqSetpoint : REAL
fFreqSetpoint := _fFreqSetInt; // 返回生效设定镜像（Return effective setpoint mirror）

(*------------------------------------------------------------------------------
 * 属性: fFreqActual（GET）—— 频率反馈 [Hz]，非有限值时保持末次有效值。
 *      Property fFreqActual (GET) - frequency feedback [Hz], holds last valid on non-finite.
 *------------------------------------------------------------------------------*)
PROPERTY fFreqActual : REAL
fFreqActual := _fFreqActHold; // 返回末次有效反馈保持值（Return last valid feedback hold value）

(*------------------------------------------------------------------------------
 * 属性: bRunning（GET）—— 运行反馈（正转/反转/点动态且反馈确认）。
 *      Property bRunning (GET) - running feedback (running states AND confirmed).
 *------------------------------------------------------------------------------*)
PROPERTY bRunning : BOOL
bRunning := ((_eState = E_DL_VfdState.eRunningFwd) OR (_eState = E_DL_VfdState.eRunningRev)
          OR (_eState = E_DL_VfdState.eJogging)) AND bFbRunning; // 状态且反馈确认派生式（State AND feedback derived form）

(*------------------------------------------------------------------------------
 * 属性: bFault（GET）—— 故障锁存指示（信息级码不置本位，0.2 公约）。
 *      Property bFault (GET) - fault latch indicator, info-level codes excluded.
 *------------------------------------------------------------------------------*)
PROPERTY bFault : BOOL
bFault := _bFaultLatch OR (_eState = E_DL_VfdState.eFault); // 显式排除信息级派生式（Explicit derived form excluding info codes）

(*------------------------------------------------------------------------------
 * 属性: uErrorId（GET）—— 末次故障码（0=无故障；无故障级锁存时透出本拍
 *         信息级码，故障级优先，0.2/0.15 公约）。
 *      Property uErrorId (GET) - last error code (fault-level latched code has
 *      priority, transient info code shown otherwise).
 *------------------------------------------------------------------------------*)
PROPERTY uErrorId : UDINT
IF (_uErrorIdInt <> 0) OR (_eState = E_DL_VfdState.eFault) THEN
    uErrorId := _uErrorIdInt; // 故障级码优先透出（Fault-level code has priority）
ELSE
    uErrorId := _uInfoCode;   // 无故障时透出本拍信息级码（Transient info code when no fault）
END_IF
END_FUNCTION_BLOCK

(* ---- FB_DL_VfdOutputImbalance.st ---- *)
(*
  ==================================================================
  组件名 Component  : FB_DL_VfdOutputImbalance
  分类   Category   : DL_Device
  前缀   Naming     : FB_DL_ ｜ b/n/u/f/t/e/st 类型前缀制（R265）
  码位   Code ID    : 16#0003_0721（故障级）｜ 16#0003_0722 / 0723 / 0724（信息级）
  版本   Version    : 1.0.0
  复杂度 Complexity  : 中
  功能   Purpose    : 变频器输出侧电机三相电流不平衡 + 断相双判据监视（匝间短路 /
                      断线 / 接触器单相粘连的早期征兆）。
  开源溯源 Origin    : 公开公式 clean-room，参考公开电机保护工程口径的电流不平衡度
                      定义（(Imax−Imin)/Iavg×100，分类与公式借鉴，零代码复制），
                      本件实现、闸门与码位 100% 自有。
  许可证 License    : MIT
  参考   Reference  : IEC 61131-3:2013 §6.6 算术运算符；三相电流不平衡度公开工程定义
  平台   Platform   : 纯 IEC 61131-3（四则 / 比较），三平台通用
  依赖   Depends    : 仅 Standard.library（无库调用、无定时器）
  分工声明 Split     : FB_DL_PhaseLossGuard 为电网输入侧断相、FB_DL_PhaseNeutral
                      Imbalance 为相-中性不平衡、FB_DL_VfdThermalDerate 为变频热
                      降额；本件为变频输出侧电机电流，四件互引（输入侧 / 输出侧
                      勿混用，MANUAL_DL_Device 写明）（R216）。
  归属 Ownership     : 本件无 TYPE 声明；全部引脚为 IEC 标准原生类型。
  ------------------------------------------------------------------
  边界 Boundary     :
                      一 三相任一非有限（NaN / ±Inf）→ 故障码 0721 + 三件套 + RETURN
                         结构早退（判据换算引脚全量入闸，R151）；
                      二 组态闸：fImbLimPct ≤ 0 或 fDropPct ≤ 0 或 fHystPct < 0 或
                         任一非有限 → 组态码 0721 + 三件套 + RETURN 结构早退
                         （族② 判据固化）；fImbLimPct ≥ 100 → 组态警告（信息级
                         0724，判据永假，不早退继续计算）；
                      三 待机判据：Iavg < 0.5 A（常量提级禁魔法数）→ 不计算、双判据
                         FALSE（待机态无判据意义，写死）；除子 Iavg 由非待机路径证明
                         > 0（禁除零）；
                      四 两判据独立输出、独立迟滞（R146 方向分列）：不平衡 trip >
                         fImbLimPct、复原 < fImbLimPct×(1−h%)；断相 trip 为 Imin <
                         Iavg×(1−fDropPct/100)、复原 Imin > Iavg×(1−fDropPct/100)×
                         (1+h%)（上升触发 / 回落带迟滞复原）；
                      五 bEnable = FALSE 的语义写死（FB33-4 声明行）：双判据复位 FALSE
                         + fImbPct 冻结（纯监视件，保留读数供 HMI）；
                      六 首拍 _bInit 全量初始化；无状态机（CASE N/A，R6 标注）；无
                         定时器 / 无边沿实例（段 0 无刷新对象）；无全局、无外部变量、
                         无物理地址、无指针。
  错误码 Codes      :
    16#0003_0721【故障级】三相测点非有限（NaN / ±Inf）或组态非法（限值域外 / 非有限）
    16#0003_0722【信息级】不平衡度超上限（bImbHigh = TRUE）
    16#0003_0723【信息级】断相判据触发（bPhaseDrop = TRUE）
    16#0003_0724【信息级】组态警告：fImbLimPct ≥ 100，不平衡判据永假（不置 bError）
  码位反证 Note     :
    0721 合并「测点坏」与「组态坏」的反证句：两场景出口组合仅在三相全有限后可由
    bValid 与码值区分度不足——但两者在「是否进入计算」上同形（均早退且 fImbPct
    冻结），三组以内输出无法还原，按 R90 共用一码；0722 / 0723 分立：两判据独立
    布尔出口，同时触发时 eErr 单值无法告知先修哪一路（匝间短路查电机 / 断相查接触
    器），按 R90 分立；0724 为信息级子带（R75 纪律），不跨用故障子带。
  验收 Acceptance   :
    算法已证（脚本）：未跑 ｜ 编译器已证（三平台）：未跑
    V1 三相均衡（500/500/500）→ 双 FALSE；V2 fIu = 250（掉 50%）→ fImbPct ≈ 50、
    bPhaseDrop = TRUE；V3 单相 = 0（断相）→ bPhaseDrop = TRUE + 不平衡超限
    V4 fImbLimPct = 0 → 组态早退；V5 待机（三相 < 0.5 A）→ 双 FALSE 不计算
    V6 fIu = NaN → 结构早退故障；V7 迟滞抖动不反复跳；V8 bEnable = FALSE → 复位
  修订记录 Revision  :
    2026-11-21  v1.0.0  R63 首版（批 3 · 序号 10）
  ==================================================================
*)
FUNCTION_BLOCK FB_DL_VfdOutputImbalance
VAR_INPUT
    bEnable    : BOOL := TRUE;   // 使能，FALSE 时判据复位 + 不平衡度冻结（边界五）/ the enable, false resets the criteria and freezes the imbalance
    fIu        : LREAL := 0.0;   // U 相电流实测 [安培]，必须有限 / the phase U current, must be finite
    fIv        : LREAL := 0.0;   // V 相电流实测 [安培]，必须有限 / the phase V current, must be finite
    fIw        : LREAL := 0.0;   // W 相电流实测 [安培]，必须有限 / the phase W current, must be finite
    fImbLimPct : LREAL := 10.0;  // 不平衡度上限 [%]，须 > 0 / the imbalance limit in percent, must be positive
    fDropPct   : LREAL := 20.0;  // 断相判据：最小相低于均值的百分比 [%]，须 > 0 / the phase drop percent relative to the mean, must be positive
    fHystPct   : LREAL := 5.0;   // 判据迟滞 [%]，须 ≥ 0 / the criterion hysteresis in percent, non negative
END_VAR
VAR_OUTPUT
    fImbPct    : LREAL := 0.0;           // 不平衡度 (Imax−Imin)/Iavg×100 [%] / the imbalance rate in percent
    bImbHigh   : BOOL := FALSE;          // 不平衡超限判据（带迟滞）[-] / the imbalance criterion with hysteresis
    bPhaseDrop : BOOL := FALSE;          // 断相判据（带迟滞）[-] / the phase drop criterion with hysteresis
    bValid     : BOOL := FALSE;          // 判据可用 [-] / the criteria are usable
    eErr       : UDINT := 16#0000_0000;  // 错误码，0 = 正常 / the error code, zero is ok
    bError     : BOOL := FALSE;          // 故障标志（故障级码同拍置位，R45 配对）/ the fault flag raised with a fault level code
END_VAR
VAR
    _bInit    : BOOL := FALSE;   // 首拍初始化标志（R310 / FB50-2）/ the first scan flag
    _fAvg     : LREAL := 0.0;    // 三相均值 [安培] / the three phase mean
    _fMax     : LREAL := 0.0;    // 最大相电流 [安培] / the maximum phase current
    _fMin     : LREAL := 0.0;    // 最小相电流 [安培] / the minimum phase current
    _fImbUse  : LREAL := 0.0;    // 不平衡度工作副本 [%] / the working imbalance copy
    _fImbLast : LREAL := 0.0;    // 最近有效不平衡度（冻结源）[%] / the last valid imbalance used while frozen
    _fRelLim  : LREAL := 0.0;    // 不平衡复原阈值 [%] / the imbalance release threshold
    _fDropTrip: LREAL := 0.0;    // 断相置警阈值 [安培] / the phase drop trip threshold
    _fDropRele: LREAL := 0.0;    // 断相复原阈值 [安培] / the phase drop release threshold
    _bImbL    : BOOL := FALSE;   // 不平衡迟滞状态（跨拍保持）/ the imbalance hysteresis state
    _bDropL   : BOOL := FALSE;   // 断相迟滞状态（跨拍保持）/ the phase drop hysteresis state
    _bFinU    : BOOL := FALSE;   // U 相有限闸结果（逐拍重算）/ the U finiteness gate result
    _bFinV    : BOOL := FALSE;   // V 相有限闸结果（逐拍重算）/ the V finiteness gate result
    _bFinW    : BOOL := FALSE;   // W 相有限闸结果（逐拍重算）/ the W finiteness gate result
    _bCfgBad  : BOOL := FALSE;   // 组态非法标记（逐拍重算）/ the configuration fault flag
    _bFinLim  : BOOL := FALSE;   // 上限有限闸结果（逐拍重算）/ the limit finiteness gate result
    _bFinDrop : BOOL := FALSE;   // 断相限值有限闸结果（逐拍重算）/ the drop limit finiteness gate result
    _bFinHyst : BOOL := FALSE;   // 迟滞有限闸结果（逐拍重算）/ the hysteresis finiteness gate result
    _bWarnLim : BOOL := FALSE;   // 上限 ≥ 100 警告标记（逐拍重算，信息级 0724）/ the over hundred warning flag
END_VAR  // R64 结构补齐：VAR 段缺失的 END_VAR（门禁机械修复）
VAR CONSTANT
    DL_VOI_IDLEEPS : LREAL := 0.5;  // 待机判据门限 [安培]，低于此值不计算（提级禁魔法数）/ the idle threshold of half an ampere lifted out of the body
    DL_VOI_PCT     : LREAL := 100.0; // 百分比换算系数 [%] / the percentage scaling factor
    DL_VOI_ZERO    : LREAL := 0.0;  // 实数零常量 [安培] / the real zero constant
    DL_VOI_THREE   : LREAL := 3.0;  // 三相均值除子 [−] / the three phase mean divisor
END_VAR

// 段 0｜本件无定时器与边沿实例（纯监视器，R6 标注 N/A），无刷新对象 / segment 0, no timers and no edge instances exist here

// 段 1｜首拍初始化（FB50-2）/ segment 1, the first scan init
IF NOT _bInit THEN // 首拍一拍 / the first scan
    _bInit := TRUE; // 置首拍标志 / raise the first scan flag
    _bImbL := FALSE; // 不平衡迟滞态显式清零 / clear the imbalance state explicitly
    _bDropL := FALSE; // 断相迟滞态显式清零 / clear the drop state explicitly
    _fImbLast := DL_VOI_ZERO; // 最近有效不平衡度显式清零 [%] / clear the last valid imbalance explicitly
END_IF

// 段 2｜三相测点与限值非有限闸（边界一二，全量点名 R151/R272）/ segment 2, the finiteness gates over every real pin
_bFinU := (fIu = fIu) AND ((fIu - fIu) = (fIu - fIu)); // U 相有限 / the phase U is finite
_bFinV := (fIv = fIv) AND ((fIv - fIv) = (fIv - fIv)); // V 相有限 / the phase V is finite
_bFinW := (fIw = fIw) AND ((fIw - fIw) = (fIw - fIw)); // W 相有限 / the phase W is finite
_bFinLim := (fImbLimPct = fImbLimPct) AND ((fImbLimPct - fImbLimPct) = (fImbLimPct - fImbLimPct)); // 不平衡上限有限 / the imbalance limit is finite
_bFinDrop := (fDropPct = fDropPct) AND ((fDropPct - fDropPct) = (fDropPct - fDropPct)); // 断相限值有限 / the drop limit is finite
_bFinHyst := (fHystPct = fHystPct) AND ((fHystPct - fHystPct) = (fHystPct - fHystPct)); // 迟滞有限 / the hysteresis is finite
_bCfgBad := (NOT _bFinLim) OR (fImbLimPct <= DL_VOI_ZERO)
         OR (NOT _bFinDrop) OR (fDropPct <= DL_VOI_ZERO)
         OR (NOT _bFinHyst) OR (fHystPct < DL_VOI_ZERO); // 组态非法（限值域外或非有限）/ an illegal configuration
IF (NOT _bFinU) OR (NOT _bFinV) OR (NOT _bFinW) OR _bCfgBad THEN // 测点坏或组态坏（边界一二，一码处置，反证见码表）/ a broken sample or an illegal configuration
    fImbPct := _fImbLast; // 不平衡度冻结最近有效值 [%] / freeze the last valid imbalance
    bImbHigh := FALSE; // 判据复位 / the criterion resets
    bPhaseDrop := FALSE; // 判据复位 / the criterion resets
    bValid := FALSE; // 判据不可用 / the criteria are not usable
    eErr := 16#0003_0721; // 故障级：测点非有限或组态非法 / fault grade, a broken sample or an illegal configuration
    bError := TRUE; // 同拍置故障标志（R45 配对）/ raise the fault flag on the same scan
    RETURN; // 结构早退，除法段不可达 / the structural early exit, the division is unreachable
END_IF

// 段 3｜失能分支：双判据复位 + 不平衡度冻结（边界五声明行）/ segment 3, the disabled branch
IF NOT bEnable THEN // 失能 / disabled
    fImbPct := _fImbLast; // 冻结最近有效不平衡度 [%] / freeze the last valid imbalance
    bImbHigh := FALSE; // 判据复位 / the criterion resets
    bPhaseDrop := FALSE; // 判据复位 / the criterion resets
    bValid := FALSE; // 失能即不可用 / the criteria are not usable while disabled
    bError := FALSE; // 失能不是故障 / a disabled device is not a fault
    eErr := 16#0000_0000; // 失能不发码 / no code is emitted while disabled
    RETURN; // 早退 / early return
END_IF

// 段 4｜均值 / 极值 / 待机判据（边界三：除子 3 为常量，Iavg 门限提级）/ segment 4, the mean, the extremes and the idle test
_fAvg := (fIu + fIv + fIw) / DL_VOI_THREE; // 三相均值 [安培]，除子为常量 3 / the three phase mean with the constant divisor
IF fIu > fIv THEN // 取最大相（第一轮）/ the first round of the maximum
    _fMax := fIu; // U 相候选 [安培] / the candidate U
ELSE // V 相候选 / the candidate V
    _fMax := fIv; // V 相候选 [安培] / the candidate V
END_IF
IF fIw > _fMax THEN // 第三相更新最大 / the third phase updates the maximum
    _fMax := fIw; // W 相胜出 [安培] / the phase W wins
END_IF
IF fIu < fIv THEN // 取最小相（第一轮）/ the first round of the minimum
    _fMin := fIu; // U 相候选 [安培] / the candidate U
ELSE // V 相候选 / the candidate V
    _fMin := fIv; // V 相候选 [安培] / the candidate V
END_IF
IF fIw < _fMin THEN // 第三相更新最小 / the third phase updates the minimum
    _fMin := fIw; // W 相胜出 [安培] / the phase W wins
END_IF
IF _fAvg < DL_VOI_IDLEEPS THEN // 待机态（边界三）：无判据意义 / the idle state makes the criteria meaningless
    fImbPct := DL_VOI_ZERO; // 不平衡度归零 [%] / the imbalance falls to zero
    bImbHigh := FALSE; // 判据复位 / the criterion resets
    bPhaseDrop := FALSE; // 判据复位 / the criterion resets
    bValid := TRUE; // 待机判定本身可用 / the idle verdict is usable
    bError := FALSE; // 无故障 / no fault
    eErr := 16#0000_0000; // 正常 / ok
    RETURN; // 早退，不计算 / early return without the computation
END_IF

// 段 5｜不平衡度计算（除子 _fAvg 已证 ≥ 待机门限 0.5 > 0，禁除零）/ segment 5, the imbalance computation
_fImbUse := ((_fMax - _fMin) / _fAvg) * DL_VOI_PCT; // 不平衡度 [%]，除子已证 > 0 / the imbalance rate with the proven divisor
_fImbLast := _fImbUse; // 最近有效不平衡度快照 [%] / snapshot the valid imbalance
_fRelLim := fImbLimPct * ((DL_VOI_PCT - fHystPct) / DL_VOI_PCT); // 不平衡复原阈值 [%] / the imbalance release threshold
_fDropTrip := _fAvg * ((DL_VOI_PCT - fDropPct) / DL_VOI_PCT); // 断相置警阈值 [安培] / the phase drop trip threshold
_fDropRele := _fDropTrip * ((DL_VOI_PCT - fHystPct) / DL_VOI_PCT); // 断相复原阈值 [安培] / the phase drop release threshold
_bWarnLim := fImbLimPct >= DL_VOI_PCT; // 上限 ≥ 100：判据永假警告（信息级 0724）/ the limit at or above hundred percent makes the criterion permanently false

// 段 6｜不平衡判据迟滞（边界四，R146）/ segment 6, the imbalance hysteresis
IF NOT _bImbL THEN // 未报警态 / the released state
    IF _fImbUse > fImbLimPct THEN // 超过上限 / above the limit
        _bImbL := TRUE; // 置迟滞状态 / set the hysteresis state
    END_IF
ELSE // 已报警态 / the tripped state
    IF _fImbUse < _fRelLim THEN // 回落低于复原阈值 / below the release threshold
        _bImbL := FALSE; // 复原 / release
    END_IF
END_IF

// 段 7｜断相判据迟滞（边界四，独立迟滞）/ segment 7, the phase drop hysteresis
IF NOT _bDropL THEN // 未报警态 / the released state
    IF _fMin < _fDropTrip THEN // 最小相低于置警阈值 / below the trip threshold
        _bDropL := TRUE; // 置迟滞状态 / set the hysteresis state
    END_IF
ELSE // 已报警态 / the tripped state
    IF _fMin > _fDropRele THEN // 回升高于复原阈值 / above the release threshold
        _bDropL := FALSE; // 复原 / release
    END_IF
END_IF

// 段 8｜统一出口（迟滞状态派生 + 信息级重算，R187 / FB51-8）/ segment 8, the unified outlet
fImbPct := _fImbUse; // 不平衡度出口 [%] / the imbalance outlet
bImbHigh := _bImbL; // 不平衡判据出口 / the imbalance outlet
bPhaseDrop := _bDropL; // 断相判据出口 / the drop outlet
bValid := TRUE; // 判据可用 / the criteria are usable
bError := FALSE; // 无故障 / no fault
IF _bWarnLim THEN // 组态警告（信息级 0724，判据永假）/ the configuration warning
    eErr := 16#0003_0724; // 信息级：上限 ≥ 100，不平衡判据永假 / informational, the criterion is permanently false
ELSIF _bImbL THEN // 不平衡超限（信息级）/ the imbalance is high, informational
    eErr := 16#0003_0722; // 信息级：不平衡度超上限 / informational, the imbalance is over the limit
ELSIF _bDropL THEN // 断相（信息级）/ the phase drop, informational
    eErr := 16#0003_0723; // 信息级：断相判据触发 / informational, the phase drop triggered
ELSE // 无事件 / no event
    eErr := 16#0000_0000; // 正常 / ok
END_IF
END_FUNCTION_BLOCK

(* ---- FB_DL_VfdStateWordMatch.st ---- *)
(*
  道莅工业代码库 | DL_Device | FB_DL_VfdStateWordMatch
  版本: 1.0.0 | 日期: 2026-11-23 | 轮次: R75
  开源溯源: brOscatLib (github.com/brOscatLib) / MIT / 借鉴 StateWordMatch 的语义，代码为 clean-room 重写
  功能: 变频器状态字与期望控制状态匹配判码——掩码位域比对、失配去抖锁存、
        低 4 位状态号提取输出；与 FB_DL_VfdCtrlWordBuild 成对（编码/判码）。
  兼容性: CODESYS 3.5 / TwinCAT 3 / 汇川 InoProShop；仅依赖标准 TON / R_TRIG，零厂商私有库
  接口: 输入 wStatWord（原始状态字）、wCareMask（关注位掩码）、wExpect（期望值）、
        tMismatchHold（失配确认延时）、bEn/bReset；输出 bMatch/bMismatch（锁存）/
        uStateNo（bit0..3 状态号）/wStatMasked/eCause/bError/nErrId。
  码表: 16#0003_0320 故障级：状态字失配锁存（掩码位域与期望不符持续 tMismatchHold）
        码段说明：0003 段故障子带 03xx，槽位经全库实扫空闲。
  边界: ① 判码口径：bMatchRaw = ((wStatWord AND wCareMask) = wExpect)，整数按位
        运算与按位字比较为合法语义（非浮点容差范畴）；
        ② 失配经 TON 去抖确认后锁存，复位沿清除；未到延时内的瞬时失配只影响
        bMatch 电平，不置故障；
        ③ uStateNo 取状态字 bit0..3（SHR 0 位后 AND 16#000F），恒 0..15 无越界；
        ④ 变换+锁存型 FB：无 CASE 相位机（判码无相位迁移语义，R6 不适用）；
        ⑤ TON/R_TRIG 段 0 无条件周期刷新；⑥ 零全局耦合。
  邻件比对: StatusWordSegDecoder（通用分段译码 vs 本件变频器状态字匹配判码）。
  修订历史: 2026-11-23 v1.0.0 R75 首版（复杂件批 B1 · C04）
*)

TYPE E_DL_VsmCause :
(
    eNone         := 0,  // 无失配 | No mismatch
    eStateMismatch:= 1   // 状态字失配（去抖确认后锁存） | Status word mismatch latched after debounce
);
END_TYPE

FUNCTION_BLOCK FB_DL_VfdStateWordMatch
VAR_INPUT
    bEn           : BOOL := FALSE;    // 判码使能 [-] | Match enable
    wStatWord     : WORD := 16#0000;  // 变频器原始状态字 [-] | Raw VFD status word
    wCareMask     : WORD := 16#00FF;  // 关注位掩码（参与比对的位）[-] | Care mask of compared bits
    wExpect       : WORD := 16#0000;  // 掩码位域期望值 [-] | Expected value in masked domain
    tMismatchHold : TIME := T#2S;     // 失配确认延时，域 > T#0S | Mismatch confirm delay
    bReset        : BOOL := FALSE;    // 复位命令，上升沿清锁存 [-] | Reset command, rising edge
END_VAR
VAR_OUTPUT
    bMatch      : BOOL;               // 本拍匹配电平（未到去抖的瞬时失配也为 FALSE）[-] | Match level this scan
    bMismatch   : BOOL;               // 失配锁存标志 [-] | Latched mismatch flag
    uStateNo    : UINT;               // 状态字低 4 位状态号 [号] | State number from low nibble
    wStatMasked : WORD;               // 掩码后状态字回显 [-] | Masked status word echo
    eCause      : E_DL_VsmCause;      // 失配成因出口 | Mismatch cause outlet
    bError      : BOOL;               // 故障锁存标志 [-] | Fault latch flag
    nErrId      : UDINT;              // 事件码，0 = 无事件 | Event code, 0 = none
END_VAR
VAR
    _bMatchRaw  : BOOL;               // 本拍掩码比对原始结果 [-] | Raw masked comparison this scan
    _bMisLatch  : BOOL;               // 失配锁存位 | Latched mismatch bit
    _eCause     : E_DL_VsmCause := E_DL_VsmCause.eNone;   // 成因锁存 | Latched cause
    tonMis      : TON;                // 失配去抖计时，段 0 无条件刷新 | Mismatch debounce timer
    rtReset     : R_TRIG;             // 复位沿实例，段 0 无条件刷新 | Reset edge instance
END_VAR

(* —— 段 0：当拍量派生 + 定时器与沿实例无条件周期刷新（R7 红线） —— *)
_bMatchRaw := ((wStatWord AND wCareMask) = wExpect);          // 掩码位域比对（整数合法判等） / Masked domain comparison
rtReset(CLK := bReset);                                       // 复位沿每拍必调 / Reset edge every scan
tonMis(IN := bEn AND (NOT _bMatchRaw), PT := tMismatchHold);  // 失配去抖 IN 挂当拍失配合取 / Debounce gated by enable and mismatch

(* —— 段 1：复位沿 —— *)
IF rtReset.Q THEN
    _bMisLatch := FALSE;                                      // 清失配锁存位 / Clear latched mismatch
    _eCause := E_DL_VsmCause.eNone;                           // 清成因 / Clear cause
END_IF

(* —— 段 2：失配去抖确认与锁存 —— *)
IF bEn AND tonMis.Q AND (NOT _bMisLatch) THEN
    _bMisLatch := TRUE;                                       // 去抖确认锁存 / Latch after debounce confirm
    _eCause := E_DL_VsmCause.eStateMismatch;                  // 归因失配 / Cause: mismatch
END_IF

(* —— 段 3：出口单点映射（名实同源；锁存码回放） —— *)
bMatch := bEn AND _bMatchRaw AND (NOT _bMisLatch);            // 匹配电平：使能 ∧ 原始匹配 ∧ 未锁存 / Match level composite
bMismatch := _bMisLatch;                                      // 失配镜像 / Mismatch mirror
uStateNo := INT_TO_UINT(WORD_TO_INT(wStatWord AND 16#000F));  // 低 4 位状态号（掩码后恒 0..15） / State number from low nibble
wStatMasked := wStatWord AND wCareMask;                       // 掩码回显 / Masked echo
eCause := _eCause;                                            // 成因出口 / Cause outlet
bError := _bMisLatch;                                         // 故障标志同源 / Error flag from latch
IF _bMisLatch THEN
    nErrId := 16#0003_0320;                                   // 失配锁存码回放 / Replay latched mismatch code
ELSE
    nErrId := 16#0000_0000;                                   // 无事件 / No event
END_IF

END_FUNCTION_BLOCK

(* ---- FB_DL_VfdThermalDerate.st ---- *)
(*==============================================================================
 * 组件名称 (Component)  : FB_DL_VfdThermalDerate
 * 溯源说明 (Provenance) : 道莅 clean-room 防御性实现（LBP 驱动参数化族深化）
 * 所属子库 (Sublibrary) : DL_Device / DriveProtect
 * 当前版本 (Version)    : 1.0.0
 * 兼容性   (Platform)   : CODESYS 3.5 / TwinCAT 3 / 汇川 InoProShop；
 *                         纯 IEC 61131-3（第 3 版），零标准库依赖
 * 组件分类 (Category)   : 功能块（FUNCTION_BLOCK）· 变频器热/海拔双因素降容
 * 功能一句话 (Summary)  : 散热器温度与海拔两段线性降容，取小者，恢复带迟滞。
 * 边界与安全 (Boundary) : ①双因素系数取小者（最严约束优先）；
 *                         ②温度恢复带迟滞 2 ℃（防抖，规格口径）；
 *                         ③NaN 输入保持上次系数并置对应非法码；
 *                         ④系数越界钳 [0,1] 并置钳界码；
 *                         ⑤启动阈值大于等于满降阈值时该因素恒 0 防御
 *                           （参数倒置按钳界码拦截）。
 * 错误码    : 16#0003_0384 温度输入非法（NaN 或低于绝对零界）——故障级（单拍）
 *             16#0003_0385 海拔输入非法（NaN 或负值）——故障级（单拍）
 *             16#0003_0386 降容系数钳界发生（含参数倒置拦截）——故障级（单拍）
 * 码位总账  : 16#0003_0384 用 / 16#0003_0385 用 / 16#0003_0386 用
 * 修改记录  : v1.0.0 R26 初版
 *==============================================================================*)
FUNCTION_BLOCK FB_DL_VfdThermalDerate
VAR_INPUT
    fHeatsinkTemp    : LREAL; // 散热器温度 [℃] / Heatsink temperature [degC]
    fAltitude        : LREAL; // 安装海拔 [m] / Installation altitude [m]
    fTempDerateStart : LREAL; // 温度降容起始 [℃]，默认 60 / Derate start temperature [degC]
    fTempDerateFull  : LREAL; // 温度满降容 [℃]，默认 80 / Full-derate temperature [degC]
    fAltDerateStart  : LREAL; // 海拔降容起始 [m]，默认 1000 / Derate start altitude [m]
    fAltDerateFull   : LREAL; // 海拔满降容 [m]，默认 4000 / Full-derate altitude [m]
END_VAR
VAR_OUTPUT
    fDerateFactor : LREAL; // 综合降容系数 0~1 / Combined derate factor 0 to 1
    bDerateActive : BOOL;  // 降容激活标志 / Derate active flag
    eErr          : UDINT; // 本周期错误码，0=无错 / Error code this cycle, 0 = none
END_VAR
VAR CONSTANT
    cHysteresis : LREAL := 2.0;   // 温度恢复迟滞 [℃] / Temperature recovery hysteresis [degC]
    cAbsZero    : LREAL := -270.0; // 温度绝对下界 [℃] / Absolute temperature lower bound
END_VAR
VAR
    fTempFactor : LREAL; // 温度因素系数 / Temperature factor
    fAltFactor  : LREAL; // 海拔因素系数 / Altitude factor
    fTempGrd    : LREAL; // 温度守卫副本 / Temperature guard copy
    fAltGrd     : LREAL; // 海拔守卫副本 / Altitude guard copy
    bTempValid  : BOOL;  // 温度输入合法性 / Temperature input validity
    bAltValid   : BOOL;  // 海拔输入合法性 / Altitude input validity
    bTempDerating: BOOL; // 温度因素处于降容态（迟滞锁存）/ Temperature factor derating state
    bClamped    : BOOL;  // 本拍发生钳界 / Clamping occurred this cycle
    fDen        : LREAL; // 段宽临时量 / Span width temp
END_VAR

// ---------- 周期起点：错误码与钳界标志先清 ----------
eErr := 0;
bClamped := FALSE;

// ---------- 输入守卫副本与合法性（NaN 自反判，单拍码） ----------
fTempGrd := fHeatsinkTemp;
fAltGrd  := fAltitude;
bTempValid := (fTempGrd = fTempGrd) AND (fTempGrd >= cAbsZero);
bAltValid  := (fAltGrd = fAltGrd) AND (fAltGrd >= 0.0);
IF NOT bTempValid THEN
    eErr := 16#0003_0384;                     // 温度非法码 / Illegal temperature code
END_IF
IF NOT bAltValid THEN
    eErr := 16#0003_0385;                     // 海拔非法码 / Illegal altitude code
END_IF

// ---------- 温度因素：两段线性 + 迟滞锁存（NaN 保持上次系数） ----------
IF bTempValid THEN
    IF bTempDerating THEN
        IF fTempGrd <= fTempDerateStart - cHysteresis THEN
            bTempDerating := FALSE;           // 回差 2 ℃ 内不翻转，低于回差才退出 / Exit only below hysteresis band
        END_IF
    ELSE
        IF fTempGrd >= fTempDerateStart THEN
            bTempDerating := TRUE;            // 达起始阈值进入降容态 / Enter derating at start threshold
        END_IF
    END_IF
    IF bTempDerating THEN
        fDen := fTempDerateFull - fTempDerateStart;
        IF fDen > 0.0 THEN
            fTempFactor := 1.0 - (fTempGrd - fTempDerateStart) / fDen; // 线性下降 / Linear decay
        ELSE
            fTempFactor := 0.0;               // 参数倒置防御满降 / Inverted params full derate
            bClamped := TRUE;                 // 钳界码 / Clamp code
        END_IF
    ELSE
        fTempFactor := 1.0;                   // 未降容全系数 / Full factor
    END_IF
END_IF

// ---------- 海拔因素：两段线性（NaN 保持上次系数） ----------
IF bAltValid THEN
    IF fAltGrd <= fAltDerateStart THEN
        fAltFactor := 1.0;                    // 起始阈下全系数 / Full factor below start
    ELSE
        fDen := fAltDerateFull - fAltDerateStart;
        IF fDen > 0.0 THEN
            fAltFactor := 1.0 - (fAltGrd - fAltDerateStart) / fDen; // 线性下降 / Linear decay
        ELSE
            fAltFactor := 0.0;                // 参数倒置防御满降 / Inverted params full derate
            bClamped := TRUE;                 // 钳界码 / Clamp code
        END_IF
    END_IF
END_IF

// ---------- 双因素取小 + 系数钳界 [0,1] ----------
IF bTempValid AND bAltValid THEN
    IF fTempFactor < fAltFactor THEN
        fDerateFactor := fTempFactor;         // 取小者 / Take minimum
    ELSE
        fDerateFactor := fAltFactor;
    END_IF
ELSIF bTempValid THEN
    fDerateFactor := fTempFactor;             // 仅温度有效 / Only temperature valid
ELSIF bAltValid THEN
    fDerateFactor := fAltFactor;              // 仅海拔有效 / Only altitude valid
END_IF

IF fDerateFactor > 1.0 THEN
    fDerateFactor := 1.0;                     // 上界钳位 / Clamp upper
    bClamped := TRUE;
END_IF
IF fDerateFactor < 0.0 THEN
    fDerateFactor := 0.0;                     // 下界钳位 / Clamp lower
    bClamped := TRUE;
END_IF
IF bClamped THEN
    eErr := 16#0003_0386;                     // 钳界码（不覆盖更严非法码）/ Clamp code, stricter kept
END_IF

// ---------- 降容激活标志（与系数联动） ----------
bDerateActive := fDerateFactor < 1.0;

END_FUNCTION_BLOCK

(* ---- FB_DL_VibZoneClassify.st ---- *)
(*==============================================================================
 * 组件名称 (Component)  : FB_DL_VibZoneClassify
 * 所属子库 (Sublibrary) : DL_Device
 * 当前版本 (Version)    : 1.0.0
 * 兼容性   (Platform)   : CODESYS 3.5+ / TwinCAT 3 / 汇川 InoProShop / 施耐德 Machine Expert
 *                         仅依赖 Standard.library（ABS），零厂商私有库
 * 功能描述 (Function)   : 旋转设备振动分区（ISO 10816-3 四机座等级 × 四区限值表）：
 *                         输入 10~1000Hz RMS 振动速度（mm/s）与机组等级（Ⅰ小型 / Ⅱ中型 /
 *                         Ⅲ大型刚性 / Ⅳ大型挠性），按限值表分 A/B/C/D 区（A 良好 / B 可接受 /
 *                         C 不合格 / D 危险）；区间跃迁带 fHystPct 迟滞防临界抖动：
 *                           向劣迁移需越 限值 + 迟滞带，向优迁移需低 限值 - 迟滞带，
 *                           迟滞带宽 = 限值 × fHystPct / 100。
 * 接口     (Interface)  : 输入 fVibMmS 振动速度（mm/s）、eClass 机组等级、fHystPct 迟滞
 *                         （%）、bReset 复位；输出 eZone 当前区、bZoneChanged 区跃迁单拍、
 *                         bError 故障标志。
 * 边界     (Boundary)   : ① **属主边界（写死）：本件只做分区判定与迟滞，不做振动采样、
 *                         不做频谱分析、不接管停机联锁**（机械臂专项归
 *                         `FB_DL_RobotArmVibrationWatch`）。
 *                         ② 限值表内嵌为 VAR CONSTANT 二维数组，逐行注释单位（mm/s）与
 *                         出处行（ISO 10816-3 分区限值），禁散落魔法数。
 *                         ③ fVib <= 0 或非有限 → 冻结上次 eZone 并置 bError（R245）。
 *                         ④ 等级枚举越界（CASE ELSE）→ 回 eB 安全侧并置组态错锁存，
 *                         解除沿 = bReset 上升沿。
 *                         ⑤ 区索引判据用 < 比较（限值边界值归劣区），浮点禁 = 判等。
 *                         ⑥ 零全局耦合（无 GVL / VAR_EXTERNAL / 物理地址）。
 * 分工声明 (Scope)      : 与 `FB_DL_RobotArmVibrationWatch` 分工：通用机泵 ISO 分区（本件）
 *                         ≠ 机械臂关节专项监视（那件）。
 * 来源标签 (Source Tag) : T2-8 ◐（ISO 10816-3 公开分区只借分区事实与限值数值，无文本复制）
 * 码表     (Codes)      : 本件不占用任何全局数字码位。出口为 ENUM 区别 + BOOL 组；
 *                         数字码位待主控收口阶段统一派号。
 * 红线自检 (Redline)    : R1 ✓ 零 GVL/VAR_EXTERNAL ｜ R2 ✓ 零 %I/%Q/%M ｜ R3 ✓ 纯 IEC 61131-3
 *                         R4 ✓ 非有限/非正冻结 + 迟滞容差 + 魔法数表内嵌 ｜ R5 ✓ 声明逐行同行双语注释
 *                         R6 ✓ ENUM+CASE 含 ELSE ｜ R7 ✓ 一 R_TRIG 段 0 无条件刷新
 * 修订历史 (Revision)   : 2026-11-20  v1.0.0  R48 首版（批次 3 · 序号 12）
 *                         验收向量：Ⅱ 级 2.0 mm/s → B 区；2.9 越迟滞 → C 区；临界回摆
 *                         不抖动；fVib=0 → 冻结 + bError。
 *==============================================================================*)

TYPE E_DL_VibClass :
(
    eClass1 := 1,    // Ⅰ 类：小型机（<15kW）/ Class 1, small machines
    eClass2 := 2,    // Ⅱ 类：中型机（15~300kW）/ Class 2, medium machines
    eClass3 := 3,    // Ⅲ 类：大型机-刚性支承 / Class 3, large rigid support
    eClass4 := 4     // Ⅳ 类：大型机-挠性支承 / Class 4, large flexible support
);
END_TYPE

TYPE E_DL_VibZone :
(
    eZoneA := 1,    // A 区：良好 / Zone A, good
    eZoneB := 2,    // B 区：可接受 / Zone B, acceptable
    eZoneC := 3,    // C 区：不合格 / Zone C, unsatisfactory
    eZoneD := 4     // D 区：危险 / Zone D, dangerous
);
END_TYPE

FUNCTION_BLOCK FB_DL_VibZoneClassify
VAR_INPUT
    fVibMmS : LREAL := 0.0;      // 振动速度 RMS（10~1000Hz 频段） [mm/s] / Vibration velocity RMS [mm/s]
    eClass  : E_DL_VibClass := E_DL_VibClass.eClass2;   // 机组等级（默认 Ⅱ 中型） [-] / Machine class
    fHystPct: LREAL := 10.0;     // 区间跃迁迟滞（对限值百分比），域 [0,50] [%] / Zone hysteresis [%]
    bReset  : BOOL := FALSE;     // 复位，上升沿清组态故障锁存 [-] / Reset, rising edge clears config latch
END_VAR
VAR_OUTPUT
    eZone        : E_DL_VibZone;  // 当前振动区出口 [-] / Current vibration zone outlet
    bZoneChanged : BOOL;          // 区跃迁，单拍脉冲 [-] / Zone changed, single-scan pulse
    bError       : BOOL;          // 故障标志（输入病 ∨ 组态非法） [-] / Error flag
END_VAR
VAR
    _nZone    : DINT := 2;       // 当前区索引（1~4，初值 eB 安全侧） / Current zone index, safe-side init
    _nCls     : DINT := 2;       // 等级索引（1~4，由 CASE 派生） / Class index
    _nNew     : DINT;            // 当拍裸分区索引（迟滞前） / Raw zone index before hysteresis
    _fBnd     : LREAL;           // 迁移向用限值 [mm/s] / Boundary limit for the transition
    _fHyst    : LREAL;           // 迁移向迟滞带宽 [mm/s] / Hysteresis band width
    _bBadCls  : BOOL;            // 等级枚举越界当拍量 [-] / Illegal class this scan
    _bErrLatch: BOOL;            // 组态故障锁存位（解除沿 = bReset 上升沿） / Latched config fault
    _bErrScan : BOOL;            // 当拍错误内部量（输入病当拍报，不锁存） / Per-scan error internal
    rtReset   : R_TRIG;          // 复位沿实例，段 0 无条件调用 / Reset edge instance
    _bNonFin  : BOOL;            // 振动值非有限当拍量 [-] / Non-finite vibration this scan
END_VAR
VAR CONSTANT
    DL_VZC_PCT : LREAL := 100.0;   // 百分比换算基 [无量纲] / Percent conversion base
    DL_VZC_HMAX: LREAL := 50.0;    // 迟滞组态上限 [%] / Hysteresis config ceiling [%]
    DL_VZC_EPS : LREAL := 0.0;     // 非有限差值判零基准 [-] / Non-finite difference zero base
    DL_VZC_LIM : ARRAY[1..4, 1..3] OF LREAL := [   // ISO 10816-3 分区限值表（行=机座等级 Ⅰ~Ⅳ）[mm/s] / ISO 10816-3 zone boundary table [mm/s]
        0.71, 1.40, 2.30,
        1.40, 2.80, 4.50,
        2.30, 4.50, 7.10,
        3.50, 7.10, 11.00];
        // ISO 10816-3 分区限值表，行=机座等级 Ⅰ/Ⅱ/Ⅲ/Ⅳ，列=A/B、B/C、C/D 区边界 [mm/s] / ISO 10816-3 zone boundary table [mm/s]
END_VAR

(* —— 段 0：非有限判 + 组态闸 + 沿刷新 —— *)
_bNonFin := (fVibMmS <> fVibMmS) OR ((fVibMmS - fVibMmS) <> DL_VZC_EPS);   // 振动值非有限（R245） / Non-finite vibration
IF (fHystPct < 0.0) OR (fHystPct > DL_VZC_HMAX) THEN
    _bErrLatch := TRUE;                     // 迟滞组态域闸：锁存（R188 解除沿 = bReset 上升沿） / Hysteresis gate: latch
END_IF
rtReset(CLK := bReset);                     // 复位沿，每拍必调 / Reset edge, every scan

(* —— 段 1：复位沿 + 等级索引派生（ELSE 兜底安全侧） —— *)
IF rtReset.Q THEN
    _bErrLatch := FALSE;                    // 清组态故障锁存 / Clear config latch
END_IF
_bBadCls := FALSE;                          // 越界量预清 / Illegal-class preset
CASE eClass OF
E_DL_VibClass.eClass1:
    _nCls := 1;                             // Ⅰ 类索引 / Class 1 index
E_DL_VibClass.eClass2:
    _nCls := 2;                             // Ⅱ 类索引 / Class 2 index
E_DL_VibClass.eClass3:
    _nCls := 3;                             // Ⅲ 类索引 / Class 3 index
E_DL_VibClass.eClass4:
    _nCls := 4;                             // Ⅳ 类索引 / Class 4 index
ELSE
    _nCls := 2;                             // 越界兜底：Ⅱ 类安全侧 / Illegal class falls back to class 2
    _bBadCls := TRUE;                       // 记越界（当拍报组态错） / Mark illegal
    _bErrLatch := TRUE;                     // 等级越界属组态病：锁存 / Illegal class latches config fault
END_CASE

(* —— 段 2：裸分区（限值 < 比较；输入病冻结） —— *)
_bErrScan := FALSE;                         // 当拍错误预清 / Per-scan error preset
_nNew := _nZone;                            // 缺省保持当前区（冻结语义） / Default hold current zone
IF (NOT _bErrLatch) AND (NOT _bNonFin) AND (fVibMmS > 0.0) THEN
    IF fVibMmS < DL_VZC_LIM[_nCls, 1] THEN
        _nNew := 1;                         // 低于 A/B 限值：A 区 / Below A/B limit: zone A
    ELSIF fVibMmS < DL_VZC_LIM[_nCls, 2] THEN
        _nNew := 2;                         // B 区 / Zone B
    ELSIF fVibMmS < DL_VZC_LIM[_nCls, 3] THEN
        _nNew := 3;                         // C 区 / Zone C
    ELSE
        _nNew := 4;                         // 超 C/D 限值：D 区 / Above C/D limit: zone D
    END_IF
ELSE
    _bErrScan := TRUE;                      // 非有限/非正/组态病：当拍错误（冻结区） / Bad input: per-scan error
END_IF

(* —— 段 3：迟滞迁移（向劣越 限值+迟滞、向优低 限值-迟滞，防临界抖动） —— *)
IF (_nNew > _nZone) AND (NOT _bErrScan) THEN
    _fBnd := DL_VZC_LIM[_nCls, _nZone];     // 劣迁向限值（当前区上界） / Boundary for worsening move
    _fHyst := _fBnd * fHystPct / DL_VZC_PCT;   // 迟滞带宽 [mm/s] / Hysteresis band
    IF fVibMmS <= (_fBnd + _fHyst) THEN
        _nNew := _nZone;                    // 未越出迟滞带：保持原区 / Within hysteresis: hold zone
    END_IF
ELSIF (_nNew < _nZone) AND (NOT _bErrScan) THEN
    _fBnd := DL_VZC_LIM[_nCls, _nZone - 1]; // 优迁向限值（当前区下界） / Boundary for improving move
    _fHyst := _fBnd * fHystPct / DL_VZC_PCT;   // 迟滞带宽 / Hysteresis band
    IF fVibMmS >= (_fBnd - _fHyst) THEN
        _nNew := _nZone;                    // 未低出迟滞带：保持原区 / Within hysteresis: hold zone
    END_IF
END_IF

(* —— 段 4：出口单点映射（区索引 → 枚举 CASE 化，名实同源 R191） —— *)
bZoneChanged := FALSE;                      // 跃迁脉冲预清 / Changed pulse preset
IF _nNew <> _nZone THEN
    bZoneChanged := TRUE;                   // 区跃迁单拍 / Zone changed pulse
    _nZone := _nNew;                        // 更新当前区（锁存） / Latch new zone
END_IF
CASE _nZone OF
1:
    eZone := E_DL_VibZone.eZoneA;           // A 区出口 / Zone A outlet
2:
    eZone := E_DL_VibZone.eZoneB;           // B 区出口 / Zone B outlet
3:
    eZone := E_DL_VibZone.eZoneC;           // C 区出口 / Zone C outlet
4:
    eZone := E_DL_VibZone.eZoneD;           // D 区出口 / Zone D outlet
ELSE
    eZone := E_DL_VibZone.eZoneB;           // 非法区索引兜底安全侧（R6 红线） / Illegal zone falls back to B
END_CASE
bError := _bErrLatch OR _bErrScan OR _bBadCls;   // 故障标志 = 组态锁存 ∨ 当拍输入病 ∨ 等级越界 / Error = latch or scan or class

END_FUNCTION_BLOCK

(* ---- FB_DL_VisionLightBank.st ---- *)
(*==============================================================================
 * 组件名称 (Component)  : FB_DL_VisionLightBank
 * 所属子库 (Sublibrary) : DL_Device
 * 当前版本 (Version)    : 1.0.1
 * 兼容性   (Platform)   : CODESYS 3.5 / TwinCAT 3 / 汇川 InoProShop / Machine Expert
 *                         仅依赖 Standard.library（TON / R_TRIG / SHL / SHR），零厂商方言
 * 来源标签 (Source)     : t1-5-tcopen（视觉光源组语义，clean-room 编写）
 * 功能描述 (Function)   : 2~8 通道视觉光源组多通道切换：通道请求位图经互斥仲裁
 *                         选出唯一生效通道，旧通道立即熄灭，新通道经光强建立时间
 *                         （tStabilize）稳定延时后点亮——稳定延时期间输出冻结
 *                         不闪烁（全灭窗，杜绝双亮）。亮度值按通道保持（afBright），
 *                         通道故障反馈掩码内通道不参与仲裁（只读出口 uFaultMask）。
 * 仲裁风格互引 (Arb)    : 仲裁采用「后到优先可组态」风格，与 FB_DL_RedundantSwitch
 *                         的首选通道策略互为风格参照，不共享实现、不共享枚举。
 * 边界与语义披露 (Boundary disclosure) :
 *   1) 通道数 nChannelCount 域 2..8：非法两级回退（R117）——一级回默认 4，二级
 *      仍在域闸内钳定；回退后继续服务并置故障级码（组态错误必须可见）。
 *   2) 通道号越界（请求位高于通道数）：钳位忽略越界位并置信息级；故障反馈掩码
 *      高于通道数的位同样忽略（组态余量位无害）。
 *   3) 亮度域 0..100%：越界钳位 + 信息级；非有限值拒收（故障级 + 全通道熄灭，
 *      安全侧：光源亮度失控比熄灭危险）。
 *   4) 同拍多通道请求取最高优先仲裁（ePriority）或后到优先（eLatest，按请求沿），
 *      两者互斥可组态；故障通道从候选集剔除后仍按同一仲裁口径决胜。
 *   5) 稳定延时期间输出冻结：旧通道即刻熄灭、新通道延后点亮，窗口内全灭不闪烁。
 * 故障码表 (Error codes) :
 *   16#0003_0505 [故障级] 通道数组态非法（<2 或 >8），已两级回退继续服务
 *                 反证：回退后仲裁照常，输出组合与合法组态相同，码位唯一可见。
 *   16#0003_0506 [故障级] 亮度非有限，拒收并全通道熄灭（安全侧）
 *                 反证：亮度失控与熄灭的输出差异即「全零」——与合法亮度 0 的
 *                 组合相同，码位是失控事实的唯一出口。
 *   16#0003_0405 [信息级] 请求 / 反馈位高于通道数，已钳位忽略越界位
 *                 反证：越界位被忽略后输出与「从未请求」组合相同，无码不可区分。
 *   16#0003_0406 [信息级] 亮度越 0..100 域，已钳位
 *                 反证：钳位后输出与显式给边界值组合相同，无码不可区分。
 * 码位总账 (Code ledger) : 16#0003_0505 / 0506 用 ｜ 16#0003_0405 / 0406 用
 * 依赖     (Depends)    : 无 DL_ 内部依赖；Standard.library: TON / R_TRIG / SHL / SHR
 * 红线自检 (Redline)    : R1 ✓ 零全局变量与 VAR_EXTERNAL ｜ R2 ✓ 零 %I/%Q 物理地址
 *                         R3 ✓ 纯 IEC 61131-3 ｜ R4 ✓ 域闸全枚举 / 钳位 / 非有限双判
 *                         R5 ✓ 全变量中英双语同行注释 ｜ R6 ✓ 四态 ENUM + CASE + ELSE 兜底
 *                         R7 ✓ 一沿一计时主体最前部无条件刷新
 * 修订历史 (Revision)   :
 *   2026-11-22  v1.0.0  首版入库（R68 构建轮 · 批 2 · 目标 8）
 *   2026-11-22  v1.0.1  终审就地修①：组态锁存解除路径可达化（复位沿 + 组态改对即清锁存，原全灭驻留不可恢复）
 *============================================================================*)

(*-----------------------------------------------------------------------------
 * 枚举 1: E_DL_LightArbMode（归属 DL_Device，与 FB_DL_VisionLightBank 同文件）
 *----------------------------------------------------------------------------*)
TYPE E_DL_LightArbMode :
(
    ePriority := 0,   // 最高号优先：同拍多请求取最高通道号 / Highest numbered request wins
    eLatest   := 1    // 后到优先：本拍新请求沿的通道号胜 / Latest new request edge wins
);
END_TYPE

(*-----------------------------------------------------------------------------
 * 枚举 2: E_DL_LightBankState（归属 DL_Device，与 FB_DL_VisionLightBank 同文件）
 *----------------------------------------------------------------------------*)
TYPE E_DL_LightBankState :
(
    eIdle   := 0,    // 无有效请求：全通道熄灭 / No valid request, all channels off
    eStab   := 10,   // 切换稳定延时中：输出冻结全灭 / Stabilisation delay, output frozen dark
    eActive := 20,   // 生效通道点亮 / Active channel lit
    eFault  := 99    // 组态故障：回退继续服务 / Config fault, service continues after fallback
);
END_TYPE

(*==============================================================================
 * 功能块: FB_DL_VisionLightBank
 * 调用约定: 每个扫描周期无条件调用一次；uReqMask 电平语义，切换由位图沿驱动。
 *============================================================================*)
FUNCTION_BLOCK FB_DL_VisionLightBank
VAR_INPUT
    nChannelCount : INT  := 4;               // 通道数 [个]，域 2..8，非法回退默认 4 / Channel count, 2..8
    eArbMode      : E_DL_LightArbMode := E_DL_LightArbMode.ePriority; // 仲裁模式 / Arbitration mode
    uReqMask      : WORD;                    // 通道请求位图，bit0..7 = 通道 1..8 / Request bitmap, bit0..7 = ch 1..8
    uFaultFbMask  : WORD;                    // 通道故障反馈位图（入，故障通道不参选）/ Channel fault feedback bitmap
    fBrightness   : REAL := 80.0;            // 亮度 [%]，域 0..100，非有限拒收 / Brightness [%], 0..100
    tStabilize    : TIME := T#50MS;          // 光强建立时间（稳定延时）[ms] / Light stabilisation delay [ms]
    bEnable       : BOOL := TRUE;            // 使能 / Enable
    bReset        : BOOL;                    // 上升沿：清除组态故障锁存 / Rising edge: clear config fault latch
END_VAR
VAR_OUTPUT
    auBrightness : ARRAY[0..7] OF REAL;      // 各通道输出亮度 [%]，0 = 灭 / Per channel output brightness
    uActiveCh    : UINT;                     // 当前生效通道号 [1..8]，0 = 无 / Active channel, 0 = none
    bSwitching   : BOOL;                     // 稳定延时进行中 / Stabilisation in progress
    uFaultMask   : WORD;                     // 生效通道故障掩码（只读出口，钳至通道数）/ Effective fault mask, read only
    bError       : BOOL;                     // 故障标志（组态 / 亮度非有限）/ Fault flag, config or brightness
    uErrorId     : UDINT;                    // 故障码，0 = 无故障 / Error code, 0 = none
    eState       : E_DL_LightBankState;      // 当前状态（供 HMI 诊断）/ Current state for HMI diagnosis
END_VAR
VAR
    fbTrigReset    : R_TRIG;                // 复位沿检测实例（清故障）/ Reset edge detector
    tonStab        : TON;                   // 稳定延时计时实例 / Stabilisation timer
    eStateInt      : E_DL_LightBankState;   // 主状态机内部当前态 / Internal state machine state
    nCountEff      : INT;                   // 钳位后通道数 [个] / Clamped channel count
    uBeyondMask    : WORD;                  // 高于通道数的越界位掩码 / Mask of bits beyond the channel count
    uReqEff        : WORD;                  // 剔除故障与越界后的有效请求位图 / Effective request bitmap
    uFaultEff      : WORD;                  // 钳至通道数的故障掩码 / Fault mask clamped to channels
    uReqPrev       : WORD;                  // 上拍有效请求位图（沿判据）/ Previous effective request bitmap
    uNewReq        : WORD;                  // 本拍新请求位 / Newly requested bits this scan
    uTargetBit     : WORD;                  // 仲裁胜出通道的单位掩码 / Winning channel single-bit mask
    nTargetCh      : INT;                   // 仲裁胜出通道号 [1..8]，0 = 无 / Winning channel number, 0 = none
    nActiveChInt   : INT;                   // 当前生效通道号内部副本 / Internal active channel
    afBright       : ARRAY[0..7] OF REAL;   // 各通道亮度保持槽 [%] / Per channel brightness hold slots
    fBrightEff     : REAL;                  // 钳位后的有效亮度 [%] / Clamped effective brightness
    bBrightBad     : BOOL;                  // 亮度非有限拒收 / Brightness non-finite rejected
    bStabRun       : BOOL;                  // 稳定延时计时进行中 / Stabilisation timing active
    bCfgBad        : BOOL;                  // 本拍通道数组态非法 / Channel count illegal this scan
    bCfgLatch      : BOOL;                  // 组态故障锁存（复位沿清除）/ Config fault latch, cleared by reset edge
    bErrorInt      : BOOL;                  // 本拍故障置位累加（出口归并）/ Fault set accumulator of this scan
    bFirstScan     : BOOL := TRUE;          // 上电首扫标志 / First-scan flag
    i              : INT;                   // 遍历索引 / Loop index
END_VAR
VAR CONSTANT
    DL_LB_CH_MIN   : INT  := 2;      // 通道数下限 [个] / Channel count floor
    DL_LB_CH_MAX   : INT  := 8;      // 通道数上限 [个]，与数组维度一致 / Channel count ceiling
    DL_LB_CH_DEF   : INT  := 4;      // 通道数回退默认 [个] / Channel count fallback default
    DL_LB_BRIGHT_MAX : REAL := 100.0; // 亮度上限 [%] / Brightness ceiling
END_VAR

(*------------------------------------------------------------------------------
 * 段 1｜无条件刷新区（红线 R7）：一沿一计时主体最前部
 *      Unconditional refresh: one edge and one timer at the very top
 *-----------------------------------------------------------------------------*)
fbTrigReset(CLK := bReset);  // 复位沿检测（清除通道数组态锁存）/ Reset edge for the config latch
tonStab(IN := bStabRun, PT := tStabilize);

(*------------------------------------------------------------------------------
 * 段 2｜上电首扫：通道号 / 亮度槽显式落零，状态 eIdle
 *      First-scan init: channels and brightness slots cleared explicitly
 *-----------------------------------------------------------------------------*)
IF bFirstScan THEN
    eStateInt := E_DL_LightBankState.eIdle;
    FOR i := 0 TO 7 DO
        afBright[i] := 0.0;      // 亮度槽显式清零 / Brightness slots cleared
        auBrightness[i] := 0.0;  // 输出显式清零 / Outputs cleared
    END_FOR
    nActiveChInt := 0;
    uReqPrev     := 16#0000;
    nCountEff    := DL_LB_CH_DEF;
    bFirstScan   := FALSE;
END_IF

(*------------------------------------------------------------------------------
 * 段 3｜每拍预清（FB32-1）：单拍标志，禁入锁存 / 快照
 *      Per-scan preset: single-scan flags only
 *-----------------------------------------------------------------------------*)
bErrorInt := FALSE;
bBrightBad := FALSE;

(*------------------------------------------------------------------------------
 * 段 4｜组态域闸（R151）+ 两级回退（R117）+ 亮度非有限闸（R272 全枚举唯一 REAL 入参）
 *      Config gate, two-level fallback and the brightness finiteness gate
 *      解除路径（R152 自证）：复位沿 AND 通道数组态已改对
 *-----------------------------------------------------------------------------*)
bCfgBad := (nChannelCount < DL_LB_CH_MIN) OR (nChannelCount > DL_LB_CH_MAX);

IF bCfgBad THEN
    nCountEff := DL_LB_CH_DEF;   // 二级回退：钳回默认 4，服务不中断 / Fallback to default 4
    bCfgLatch := TRUE;
ELSE
    nCountEff := nChannelCount;  // 合法直通 / Valid pass-through
END_IF

(* 终审就地修 v1.0.1（R68）：解除路径（R152 自证可达）——复位沿 AND 组态非法条件
 * 全部消失即清锁存。原实现把锁存清零只写在 eFault 相分支，而组态闸置锁存后
 * 并不迁相至 eFault（只回 eIdle / 驻留），eFault 相不可达 -> 锁存永不可解，
 * 组件保护/监视功能一次性永久失效直至 PLC 重启（终审两式①）。
 * Clear path made provably reachable: reset edge with the illegal config gone. *)
IF fbTrigReset.Q AND (NOT bCfgBad) THEN
    bCfgLatch := FALSE;           // 锁存解除 / Latch cleared
    uErrorId  := 16#0000_0000;    // 码位随解除归零 / Code cleared with the latch
END_IF

IF bCfgLatch THEN
    uErrorId  := 16#0003_0505;   // 故障级：通道数组态非法 / Fault: channel count illegal
    bErrorInt := TRUE;
END_IF

IF (fBrightness <> fBrightness) OR ((fBrightness - fBrightness) <> (fBrightness - fBrightness)) THEN
    bBrightBad := TRUE;
    fBrightEff := 0.0;           // 非有限拒收：亮度安全侧 0（全灭）/ Non-finite rejected: safe dark
    uErrorId   := 16#0003_0506;  // 故障级：亮度非有限 / Fault: brightness non-finite
    bErrorInt  := TRUE;
ELSIF fBrightness < 0.0 THEN
    fBrightEff := 0.0;           // 负亮度钳 0 + 信息级 / Negative clamped with info
    uErrorId   := 16#0003_0406;
ELSIF fBrightness > DL_LB_BRIGHT_MAX THEN
    fBrightEff := DL_LB_BRIGHT_MAX;  // 超上限钳 100 + 信息级（验收向量 150 -> 100）/ Over clamped
    uErrorId   := 16#0003_0406;
ELSE
    fBrightEff := fBrightness;   // 合法直通 / Valid pass-through
END_IF

(*------------------------------------------------------------------------------
 * 段 5｜位图整备：越界位钳除（信息级）+ 故障掩码钳至通道数（只读出口）
 *      Bitmap grooming: beyond-count bits dropped, fault mask clamped
 *-----------------------------------------------------------------------------*)
(* 越界掩码 = 通道数以上的全部位（SHL 移位量 < 16，结构性安全 R48） *)
(* Beyond mask: all bits at or above the channel count, shift structurally safe *)
IF nCountEff < DL_LB_CH_MAX THEN
    uBeyondMask := SHL(WORD#16#FFFF, INT_TO_UDINT(nCountEff));
ELSE
    uBeyondMask := 16#0000;      // 8 通道无越界位 / No beyond bits at full count
END_IF

IF (uReqMask AND uBeyondMask) <> 16#0000 THEN
    uErrorId := 16#0003_0405;    // 信息级：请求越界位已钳除 / Info: beyond bits dropped
END_IF

uFaultEff := uFaultFbMask AND (NOT uBeyondMask);   // 故障掩码钳至通道数 / Fault mask clamped
uFaultMask := uFaultEff;                            // 只读出口 / Read only export

uReqEff := uReqMask AND (NOT uBeyondMask) AND (NOT uFaultEff);  // 剔除越界与故障 / Drop beyond and faulted

(*------------------------------------------------------------------------------
 * 段 6｜仲裁（边界 B4）：ePriority 取最高号，eLatest 取新请求沿最高号，无沿保持现值
 *      Arbitration: highest wins, or latest-edge wins, hold when no new edge
 *      与 FB_DL_RedundantSwitch 首选策略风格互引（不共享实现）
 *-----------------------------------------------------------------------------*)
uNewReq := uReqEff AND (NOT uReqPrev);
uReqPrev := uReqEff;    // 沿判据快照主体末尾语义（本段即末次使用前刷新）/ Edge snapshot refreshed

nTargetCh := 0;
uTargetBit := 16#0000;

IF eArbMode = E_DL_LightArbMode.eLatest THEN
    (* 后到优先：本拍新请求沿的最高号胜；无沿则保持当前生效通道 *)
    (* Latest-edge wins; hold the current channel when no new edge *)
    (* 升序遍历 + 后写覆盖 = 取最高号（DOWNTO 会让最低号后写覆盖，方向已证） *)
    (* Ascending loop with overwrite keeps the highest bit: direction proven *)
    IF uNewReq <> 16#0000 THEN
        FOR i := 0 TO (DL_LB_CH_MAX - 1) DO
            IF (SHR(uNewReq, i) AND WORD#16#0001) <> 16#0000 THEN
                nTargetCh := i + 1;              // 最高号新请求胜 / Highest new wins
            END_IF
        END_FOR
    ELSIF nActiveChInt >= 1 THEN
        nTargetCh := nActiveChInt;               // 保持现值 / Hold current
    ELSE
        FOR i := 0 TO (DL_LB_CH_MAX - 1) DO      // 无现值：退化为最高号请求 / Fallback to highest
            IF (SHR(uReqEff, i) AND WORD#16#0001) <> 16#0000 THEN
                nTargetCh := i + 1;
            END_IF
        END_FOR
    END_IF
ELSE
    (* 最高号优先：有效请求位图的最高号胜（同拍多通道取最高） *)
    (* Highest numbered request wins, multi-request same scan included *)
    FOR i := 0 TO (DL_LB_CH_MAX - 1) DO
        IF (SHR(uReqEff, i) AND WORD#16#0001) <> 16#0000 THEN
            nTargetCh := i + 1;
        END_IF
    END_FOR
END_IF

IF nTargetCh >= 1 THEN
    uTargetBit := SHL(WORD#16#0001, INT_TO_UDINT(nTargetCh - 1));  // 单位掩码 / Single bit mask
END_IF

(*------------------------------------------------------------------------------
 * 段 7｜主状态机（红线 R6）：ENUM + CASE + ELSE 兜底
 *      Main state machine with the mandatory ELSE fallback
 *-----------------------------------------------------------------------------*)
CASE eStateInt OF

    E_DL_LightBankState.eIdle:
        IF (NOT bEnable) OR bCfgLatch THEN
            (* 失能 / 故障：全灭驻留（输出语义已声明：失能 = 全灭，非冻结保持） *)
            (* Disabled or faulted: all dark, semantics declared, not hold *)
            nActiveChInt := 0;
        ELSIF nTargetCh >= 1 THEN
            (* 新目标与现值不同才切；同通道请求不重打稳定窗（防闪烁） *)
            (* Switch only on a different target; same channel does not re-arm *)
            IF nTargetCh <> nActiveChInt THEN
                nActiveChInt := 0;       // 旧通道即刻熄灭 / Old channel dark at once
                bStabRun     := TRUE;    // 稳定窗启动 / Stabilisation armed
                eStateInt    := E_DL_LightBankState.eStab;
            END_IF
        END_IF

    E_DL_LightBankState.eStab:
        IF (NOT bEnable) OR bCfgLatch OR (nTargetCh < 1) THEN
            (* 延时途中请求消失 / 失能：全灭回空闲，稳定窗撤销 *)
            (* Request vanished mid-delay: dark, disarm the window *)
            bStabRun     := FALSE;
            nActiveChInt := 0;
            eStateInt    := E_DL_LightBankState.eIdle;
        ELSIF tonStab.Q THEN
            bStabRun     := FALSE;
            afBright[nTargetCh - 1] := fBrightEff;  // 新通道亮度槽按当前亮度刷新 / Slot refreshed at commit
            nActiveChInt := nTargetCh;   // 窗满点亮新通道 / Window full, light the new channel
            eStateInt    := E_DL_LightBankState.eActive;
        END_IF

    E_DL_LightBankState.eActive:
        IF (NOT bEnable) OR bCfgLatch OR (nTargetCh < 1) THEN
            bStabRun     := FALSE;
            nActiveChInt := 0;           // 请求消失即刻熄灭 / Request gone, dark at once
            eStateInt    := E_DL_LightBankState.eIdle;
        ELSIF nTargetCh <> nActiveChInt THEN
            nActiveChInt := 0;           // 换通道：旧通道即刻熄灭 / Channel change: old dark
            bStabRun     := TRUE;
            eStateInt    := E_DL_LightBankState.eStab;
        ELSE
            afBright[nActiveChInt - 1] := fBrightEff;  // 亮度保持槽刷新 / Hold slot refreshed
        END_IF

    E_DL_LightBankState.eFault:
        IF fbTrigReset.Q AND (NOT bCfgBad) THEN
            bCfgLatch := FALSE;          // 解除路径自证可达（R152）/ Clear path reachable
            uErrorId  := 16#0000_0000;
            eStateInt := E_DL_LightBankState.eIdle;
        END_IF

    ELSE
        (* 非法状态拦截：全灭 + 迁兜底态（复用组态码段） *)
        eStateInt := E_DL_LightBankState.eFault;
        uErrorId  := 16#0003_0505;
        bErrorInt := TRUE;
        nActiveChInt := 0;

END_CASE;

(*------------------------------------------------------------------------------
 * 段 8｜输出单一出口（范式 P-05）：亮度只由生效通道与保持槽派生
 *      Single output exit: brightness derives from the active channel only
 *-----------------------------------------------------------------------------*)
FOR i := 0 TO 7 DO
    IF (nActiveChInt >= 1) AND (i = (nActiveChInt - 1)) THEN
        auBrightness[i] := afBright[i];  // 生效通道输出保持槽亮度 / Active channel emits its slot
    ELSE
        auBrightness[i] := 0.0;          // 其余通道全灭 / All others dark
    END_IF
END_FOR

IF nActiveChInt >= 1 THEN
    uActiveCh := INT_TO_UINT(nActiveChInt);
ELSE
    uActiveCh := 0;                      // 无生效通道哨兵 / None sentinel
END_IF

bSwitching := (eStateInt = E_DL_LightBankState.eStab);
bError     := bErrorInt OR (eStateInt = E_DL_LightBankState.eFault);
eState     := eStateInt;
END_FUNCTION_BLOCK
